(* IEC 61131-3 sources: plc-st-coding-agent/progress/evidence/f14_v14_remaining_20261113/jobs/codex_minimax-m27 (part 4) *)

(* ---- public-medium-04.patch_base_04.st ---- *)
FUNCTION_BLOCK FB_TemperatureControl
VAR_INPUT
    TemperatureSensorInput : REAL;
    SetTemperature : REAL;
END_VAR

VAR_OUTPUT
    CurrentTemperature : REAL;
    SetTempDisplay : REAL;
    HeaterStatus : BOOL;
    OverheatProtection : BOOL;
    HeaterOutput : BOOL;
END_VAR

VAR
    HeaterRuntimeTimer : TON;
    OverheatCooldownTimer : TON;
    tmp_InOverheatProtection : BOOL;
    tmp_SensorFault : BOOL;
    tmp_HeaterShouldBeOn : BOOL;
END_VAR

(*
ENGINEERING_CONTRACT
================================================================================
| Output/State        | Activation          | Retention/Reset           | Units/Boundaries     |
|---------------------|---------------------|---------------------------|----------------------|
| CurrentTemperature  | Every scan (copy)   | Unchanged when fault      | REAL, no conversion  |
| SetTempDisplay      | Every scan (copy)   | Always updated            | REAL, no conversion  |
| HeaterStatus        | Every scan (AND)    | False on fault or overheat| BOOL, same-scan      |
| OverheatProtection  | tmp_InOverheatProt  | Hold 3s cooldown then OFF | BOOL, timer-driven   |
| HeaterOutput        | temp < set && !prot | Off on fault, >5s prot,   | BOOL, 5s threshold   |
|                     |                     |   or temp >= set          | > not >= per spec    |
================================================================================
PUB001: temp < set triggers heater on
PUB002: temp > set turns heater off
PUB003: >5s continuous heater runtime triggers overheat protection
PUB004: 3s cooldown before overheat protection can be lifted
PUB005: Sensor fault if input < 0 or > 100
PUB006: Display current temp, set temp, heater status, overheat status
PUB007: Heater must be off during sensor fault
PUB008: Heater off during overheat protection until cooldown completes
================================================================================

CONTRACT_RULES []
*)

// Update display outputs every scan
CurrentTemperature := TemperatureSensorInput;
SetTempDisplay := SetTemperature;

// Detect sensor fault: temperature out of valid range [0, 100]
tmp_SensorFault := (TemperatureSensorInput < 0.0) OR (TemperatureSensorInput > 100.0);

// Determine if heater should be on (based on temperature comparison only)
tmp_HeaterShouldBeOn := (NOT tmp_SensorFault) AND (TemperatureSensorInput < SetTemperature);

// Overheat protection state machine
IF NOT tmp_InOverheatProtection THEN
    // Normal operation: check if overheat protection should trigger
    IF tmp_HeaterShouldBeOn THEN
        // Heater is on, start accumulating runtime
        HeaterRuntimeTimer(IN := TRUE, PT := T#5S);
        IF HeaterRuntimeTimer.Q THEN
            // Heater ran for more than 5 seconds continuously
            tmp_InOverheatProtection := TRUE;
            HeaterRuntimeTimer(IN := FALSE);
        END_IF;
    ELSE
        // Heater is off, reset runtime timer
        HeaterRuntimeTimer(IN := FALSE);
    END_IF;
ELSE
    // In overheat protection state, start 3-second cooldown
    HeaterRuntimeTimer(IN := FALSE);
    OverheatCooldownTimer(IN := TRUE, PT := T#3S);
    IF OverheatCooldownTimer.Q THEN
        // Cooldown complete, clear overheat protection
        tmp_InOverheatProtection := FALSE;
        OverheatCooldownTimer(IN := FALSE);
    END_IF;
END_IF;

// Update overheat protection output
OverheatProtection := tmp_InOverheatProtection;

// Calculate final heater output
// HeaterOutput is true when:
//   - Temperature is below setpoint
//   - Not in sensor fault
//   - Not in overheat protection
HeaterOutput := tmp_HeaterShouldBeOn AND (NOT tmp_InOverheatProtection);

// Heater status follows actual heater output
HeaterStatus := HeaterOutput;

END_FUNCTION_BLOCK

(* ---- public-medium-04.raw_candidate_01.st ---- *)
FUNCTION_BLOCK FB_TemperatureControl
VAR_INPUT
    TemperatureSensorInput : REAL;
    SetTemperature : REAL;
END_VAR

VAR_OUTPUT
    CurrentTemperature : REAL;
    SetTempDisplay : REAL;
    HeaterStatus : BOOL;
    OverheatProtection : BOOL;
    HeaterOutput : BOOL;
END_VAR

VAR
    HeaterRuntimeTimer : TON;
    OverheatCooldownTimer : TON;
    tmp_InOverheatProtection : BOOL;
    tmp_SensorFault : BOOL;
END_VAR

(*
ENGINEERING_CONTRACT
================================================================================
| Output/State        | Activation          | Retention/Reset           | Units/Boundaries     |
|---------------------|---------------------|---------------------------|----------------------|
| CurrentTemperature  | Every scan (copy)   | Unchanged when fault      | REAL, no conversion  |
| SetTempDisplay      | Every scan (copy)   | Always updated            | REAL, no conversion  |
| HeaterStatus        | Every scan (AND)    | False on fault or overheat| BOOL, same-scan      |
| OverheatProtection  | tmp_InOverheatProt  | Hold 3s cooldown then OFF | BOOL, timer-driven   |
| HeaterOutput        | temp < set && !prot | Off on fault, >5s prot,   | BOOL, 5s threshold   |
|                     |                     |   or temp >= set          | > not >= per spec    |
================================================================================
PUB001: temp < set triggers heater on
PUB002: temp > set turns heater off
PUB003: >5s continuous heater runtime triggers overheat protection
PUB004: 3s cooldown before overheat protection can be lifted
PUB005: Sensor fault if input < 0 or > 100
PUB006: Display current temp, set temp, heater status, overheat status
PUB007: Heater must be off during sensor fault
PUB008: Heater off during overheat protection until cooldown completes
================================================================================

CONTRACT_RULES []
*)

// Update display outputs every scan
CurrentTemperature := TemperatureSensorInput;
SetTempDisplay := SetTemperature;

// Detect sensor fault: temperature out of valid range [0, 100]
tmp_SensorFault := (TemperatureSensorInput < 0.0) OR (TemperatureSensorInput > 100.0);

// Determine if heater should be on (based on temperature comparison only)
tmp_HeaterShouldBeOn := (NOT tmp_SensorFault) AND (TemperatureSensorInput < SetTemperature);

// Overheat protection state machine
IF NOT tmp_InOverheatProtection THEN
    // Normal operation: check if overheat protection should trigger
    IF tmp_HeaterShouldBeOn THEN
        // Heater is on, start accumulating runtime
        HeaterRuntimeTimer(IN := TRUE, PT := T#5S);
        IF HeaterRuntimeTimer.Q THEN
            // Heater ran for more than 5 seconds continuously
            tmp_InOverheatProtection := TRUE;
            HeaterRuntimeTimer(IN := FALSE);
        END_IF;
    ELSE
        // Heater is off, reset runtime timer
        HeaterRuntimeTimer(IN := FALSE);
    END_IF;
ELSE
    // In overheat protection state, start 3-second cooldown
    HeaterRuntimeTimer(IN := FALSE);
    OverheatCooldownTimer(IN := TRUE, PT := T#3S);
    IF OverheatCooldownTimer.Q THEN
        // Cooldown complete, clear overheat protection
        tmp_InOverheatProtection := FALSE;
        OverheatCooldownTimer(IN := FALSE);
    END_IF;
END_IF;

// Update overheat protection output
OverheatProtection := tmp_InOverheatProtection;

// Calculate final heater output
// HeaterOutput is true when:
//   - Temperature is below setpoint
//   - Not in sensor fault
//   - Not in overheat protection
HeaterOutput := tmp_HeaterShouldBeOn AND (NOT tmp_InOverheatProtection);

// Heater status follows actual heater output
HeaterStatus := HeaterOutput;

END_FUNCTION_BLOCK

(* ---- public-medium-04.raw_candidate_02.st ---- *)
FUNCTION_BLOCK FB_TemperatureControl
VAR_INPUT
    TemperatureSensorInput : REAL;
    SetTemperature : REAL;
END_VAR

VAR_OUTPUT
    CurrentTemperature : REAL;
    SetTempDisplay : REAL;
    HeaterStatus : BOOL;
    OverheatProtection : BOOL;
    HeaterOutput : BOOL;
END_VAR

VAR
    HeaterRuntimeTimer : TON;
    OverheatCooldownTimer : TON;
    tmp_InOverheatProtection : BOOL;
    tmp_SensorFault : BOOL;
    tmp_HeaterShouldBeOn : BOOL;
END_VAR

(*
ENGINEERING_CONTRACT
================================================================================
| Output/State        | Activation          | Retention/Reset           | Units/Boundaries     |
|---------------------|---------------------|---------------------------|----------------------|
| CurrentTemperature  | Every scan (copy)   | Unchanged when fault      | REAL, no conversion  |
| SetTempDisplay      | Every scan (copy)   | Always updated            | REAL, no conversion  |
| HeaterStatus        | Every scan (AND)    | False on fault or overheat| BOOL, same-scan      |
| OverheatProtection  | tmp_InOverheatProt  | Hold 3s cooldown then OFF | BOOL, timer-driven   |
| HeaterOutput        | temp < set && !prot | Off on fault, >5s prot,   | BOOL, 5s threshold   |
|                     |                     |   or temp >= set          | > not >= per spec    |
================================================================================
PUB001: temp < set triggers heater on
PUB002: temp > set turns heater off
PUB003: >5s continuous heater runtime triggers overheat protection
PUB004: 3s cooldown before overheat protection can be lifted
PUB005: Sensor fault if input < 0 or > 100
PUB006: Display current temp, set temp, heater status, overheat status
PUB007: Heater must be off during sensor fault
PUB008: Heater off during overheat protection until cooldown completes
================================================================================

CONTRACT_RULES []
*)

// Update display outputs every scan
CurrentTemperature := TemperatureSensorInput;
SetTempDisplay := SetTemperature;

// Detect sensor fault: temperature out of valid range [0, 100]
tmp_SensorFault := (TemperatureSensorInput < 0.0) OR (TemperatureSensorInput > 100.0);

// Determine if heater should be on (based on temperature comparison only)
tmp_HeaterShouldBeOn := (NOT tmp_SensorFault) AND (TemperatureSensorInput < SetTemperature);

// Overheat protection state machine
IF NOT tmp_InOverheatProtection THEN
    // Normal operation: check if overheat protection should trigger
    IF tmp_HeaterShouldBeOn THEN
        // Heater is on, start accumulating runtime
        HeaterRuntimeTimer(IN := TRUE, PT := T#5S);
        IF HeaterRuntimeTimer.Q THEN
            // Heater ran for more than 5 seconds continuously
            tmp_InOverheatProtection := TRUE;
            HeaterRuntimeTimer(IN := FALSE);
        END_IF;
    ELSE
        // Heater is off, reset runtime timer
        HeaterRuntimeTimer(IN := FALSE);
    END_IF;
ELSE
    // In overheat protection state, start 3-second cooldown
    HeaterRuntimeTimer(IN := FALSE);
    OverheatCooldownTimer(IN := TRUE, PT := T#3S);
    IF OverheatCooldownTimer.Q THEN
        // Cooldown complete, clear overheat protection
        tmp_InOverheatProtection := FALSE;
        OverheatCooldownTimer(IN := FALSE);
    END_IF;
END_IF;

// Update overheat protection output
OverheatProtection := tmp_InOverheatProtection;

// Calculate final heater output
// HeaterOutput is true when:
//   - Temperature is below setpoint
//   - Not in sensor fault
//   - Not in overheat protection
HeaterOutput := tmp_HeaterShouldBeOn AND (NOT tmp_InOverheatProtection);

// Heater status follows actual heater output
HeaterStatus := HeaterOutput;

END_FUNCTION_BLOCK

(* ---- public-medium-04.raw_candidate_04.st ---- *)
FUNCTION_BLOCK FB_TemperatureControl
VAR_INPUT
    TemperatureSensorInput : REAL;
    SetTemperature : REAL;
END_VAR

VAR_OUTPUT
    CurrentTemperature : REAL;
    SetTempDisplay : REAL;
    HeaterStatus : BOOL;
    OverheatProtection : BOOL;
    HeaterOutput : BOOL;
END_VAR

VAR
    HeaterRuntimeTimer : TON;
    OverheatCooldownTimer : TON;
    tmp_InOverheatProtection : BOOL;
    tmp_SensorFault : BOOL;
    tmp_RuntimeTimerEnable : BOOL;
END_VAR

(*
ENGINEERING_CONTRACT
================================================================================
| Output/State        | Activation          | Retention/Reset           | Units/Boundaries     |
|---------------------|---------------------|---------------------------|----------------------|
| CurrentTemperature  | Every scan (copy)   | Unchanged when fault      | REAL, no conversion  |
| SetTempDisplay      | Every scan (copy)   | Always updated            | REAL, no conversion  |
| HeaterStatus        | Every scan (AND)    | False on fault or overheat| BOOL, same-scan      |
| OverheatProtection  | tmp_InOverheatProt  | Hold 3s cooldown then OFF | BOOL, timer-driven   |
| HeaterOutput        | temp < set && !prot | Off on fault, >5s prot,   | BOOL, 5s threshold   |
|                     |                     |   or temp >= set          | > not >= per spec    |
================================================================================
PUB001: temp < set triggers heater on
PUB002: temp > set turns heater off
PUB003: >5s continuous heater runtime triggers overheat protection
PUB004: 3s cooldown before overheat protection can be lifted
PUB005: Sensor fault if input < 0 or > 100
PUB006: Display current temp, set temp, heater status, overheat status
PUB007: Heater must be off during sensor fault
PUB008: Heater off during overheat protection until cooldown completes
================================================================================

CONTRACT_RULES []
*)

// Update display outputs every scan
CurrentTemperature := TemperatureSensorInput;
SetTempDisplay := SetTemperature;

// Detect sensor fault: temperature out of valid range [0, 100]
tmp_SensorFault := (TemperatureSensorInput < 0.0) OR (TemperatureSensorInput > 100.0);

// Determine if runtime timer should accumulate (heater on, not in fault, not in overheat protection)
tmp_RuntimeTimerEnable := (NOT tmp_SensorFault) AND (NOT tmp_InOverheatProtection) AND (TemperatureSensorInput < SetTemperature);

// Overheat protection state machine
IF NOT tmp_InOverheatProtection THEN
    // Normal operation: check if overheat protection should trigger
    IF tmp_RuntimeTimerEnable THEN
        // Heater is on, start accumulating runtime
        HeaterRuntimeTimer(IN := TRUE, PT := T#5001MS);
        IF HeaterRuntimeTimer.Q THEN
            // Heater ran for more than 5 seconds continuously
            tmp_InOverheatProtection := TRUE;
            HeaterRuntimeTimer(IN := FALSE);
        END_IF;
    ELSE
        // Heater is off or in fault, reset runtime timer
        HeaterRuntimeTimer(IN := FALSE);
    END_IF;
ELSE
    // In overheat protection state, run 3-second cooldown
    HeaterRuntimeTimer(IN := FALSE);
    OverheatCooldownTimer(IN := TRUE, PT := T#3S);
    IF OverheatCooldownTimer.Q THEN
        // Cooldown complete, clear overheat protection
        tmp_InOverheatProtection := FALSE;
        OverheatCooldownTimer(IN := FALSE);
    END_IF;
END_IF;

// Update outputs
OverheatProtection := tmp_InOverheatProtection;

// Calculate final heater output: on when temperature below setpoint, not in fault, not in overheat protection
HeaterOutput := tmp_RuntimeTimerEnable;

// Heater status follows actual heater output
HeaterStatus := HeaterOutput;

END_FUNCTION_BLOCK

(* ---- public-medium-05.candidate_01.st ---- *)
(* ENGINEERING_CONTRACT *)
(*
Mode behavior (PUB001):
- Mode=0: Manual mode (ForwardButton→MotorForward, ReverseButton→MotorReverse)
- Mode=1: Automatic mode (A→B→C state machine)

Manual mode (PUB002):
- MotorForward activates with ForwardButton when Mode=0, interlocked with ReverseButton
- MotorReverse activates with ReverseButton when Mode=0, interlocked with ForwardButton
- CompletionLight always OFF in manual mode

Automatic mode (PUB003):
- IDLE→SensorA: wait at Station A for ButtonA press
- Station A: MotorForward TRUE while State=MOVING_TO_B
- MOVING_TO_B→SensorB: hold at Station B for ButtonB press
- Station B: MotorForward TRUE while State=MOVING_TO_C
- MOVING_TO_C→SensorC: hold at Station C

CompletionLight behavior (PUB006, PUB007, PUB008):
- Activation: State=STATION_C AND SensorC AND ButtonC (same-scan)
- Retention: State=STATION_C AND SensorC (CompletionLight remains TRUE)
- Deactivation: State≠STATION_C OR NOT SensorC (product removal)
- Units: boolean, no units

Output states:
- MotorForward: combinational in manual, pulsed in auto (A→B, B→C transitions)
- MotorReverse: combinational in manual only, always FALSE in auto
- CompletionLight: retained while product at Station C, no explicit reset input

Scan priority: same-scan evaluation of all conditions before outputs
*)

(* CONTRACT_RULES [] *)

FUNCTION_BLOCK ProductionLineControl
VAR_INPUT
    Mode            : BOOL;
    ForwardButton   : BOOL;
    ReverseButton   : BOOL;
    SensorA         : BOOL;
    SensorB         : BOOL;
    SensorC         : BOOL;
    ButtonA         : BOOL;
    ButtonB         : BOOL;
    ButtonC         : BOOL;
END_VAR
VAR_OUTPUT
    MotorForward    : BOOL;
    MotorReverse    : BOOL;
    CompletionLight : BOOL;
END_VAR
VAR
    State : INT;
END_VAR

// State constants
CONSTANTS
    STATE_IDLE         : INT := 0;
    STATE_STATION_A    : INT := 1;
    STATE_MOVING_TO_B  : INT := 2;
    STATE_STATION_B    : INT := 3;
    STATE_MOVING_TO_C  : INT := 4;
    STATE_STATION_C    : INT := 5;
END_CONSTANTS

// Initialize state on first call
IF State = 0 THEN
    State := STATE_IDLE;
END_IF;

// Manual mode: direct button control with direction interlock
IF Mode = FALSE THEN
    MotorForward := ForwardButton AND NOT ReverseButton;
    MotorReverse := ReverseButton AND NOT ForwardButton;
    CompletionLight := FALSE;
    State := STATE_IDLE;
ELSE
    // Automatic mode: state machine control
    IF State = STATE_IDLE THEN
        MotorForward := FALSE;
        MotorReverse := FALSE;
        CompletionLight := FALSE;

        IF SensorA THEN
            State := STATE_STATION_A;
        END_IF;

    ELSIF State = STATE_STATION_A THEN
        MotorForward := FALSE;

        IF ButtonA THEN
            State := STATE_MOVING_TO_B;
        END_IF;

    ELSIF State = STATE_MOVING_TO_B THEN
        MotorForward := TRUE;

        IF SensorB THEN
            MotorForward := FALSE;
            State := STATE_STATION_B;
        END_IF;

    ELSIF State = STATE_STATION_B THEN
        MotorForward := FALSE;

        IF ButtonB THEN
            State := STATE_MOVING_TO_C;
        END_IF;

    ELSIF State = STATE_MOVING_TO_C THEN
        MotorForward := TRUE;

        IF SensorC THEN
            MotorForward := FALSE;
            State := STATE_STATION_C;
        END_IF;

    ELSIF State = STATE_STATION_C THEN
        MotorForward := FALSE;

        IF NOT SensorC THEN
            State := STATE_IDLE;
            CompletionLight := FALSE;
        ELSE
            CompletionLight := TRUE;
        END_IF;
    END_IF;
END_IF;

END_FUNCTION_BLOCK

(* ---- public-medium-05.patch_base_02.st ---- *)
(* ENGINEERING_CONTRACT *)
(*
Mode behavior (PUB001):
- Mode=0: Manual mode (ForwardButton→MotorForward, ReverseButton→MotorReverse)
- Mode=1: Automatic mode (A→B→C state machine)

Manual mode (PUB002):
- MotorForward activates with ForwardButton when Mode=0, interlocked with ReverseButton
- MotorReverse activates with ReverseButton when Mode=0, interlocked with ForwardButton
- CompletionLight always OFF in manual mode

Automatic mode (PUB003):
- IDLE→SensorA: wait at Station A for ButtonA press
- Station A: MotorForward TRUE while State=MOVING_TO_B
- MOVING_TO_B→SensorB: hold at Station B for ButtonB press
- Station B: MotorForward TRUE while State=MOVING_TO_C
- MOVING_TO_C→SensorC: hold at Station C

CompletionLight behavior (PUB006, PUB007, PUB008):
- Activation: State=STATION_C AND SensorC AND ButtonC (same-scan)
- Retention: State=STATION_C AND SensorC (CompletionLight remains TRUE)
- Deactivation: State≠STATION_C OR NOT SensorC (product removal)
- Units: boolean, no units

Output states:
- MotorForward: combinational in manual, pulsed in auto (A→B, B→C transitions)
- MotorReverse: combinational in manual only, always FALSE in auto
- CompletionLight: retained while product at Station C, no explicit reset input

Scan priority: same-scan evaluation of all conditions before outputs
*)

(* CONTRACT_RULES [] *)

FUNCTION_BLOCK ProductionLineControl
VAR_INPUT
    Mode            : BOOL;
    ForwardButton   : BOOL;
    ReverseButton   : BOOL;
    SensorA         : BOOL;
    SensorB         : BOOL;
    SensorC         : BOOL;
    ButtonA         : BOOL;
    ButtonB         : BOOL;
    ButtonC         : BOOL;
END_VAR
VAR_OUTPUT
    MotorForward    : BOOL;
    MotorReverse    : BOOL;
    CompletionLight : BOOL;
END_VAR
VAR
    State : INT;
END_VAR

// State constants
CONSTANTS
    STATE_IDLE         : INT := 0;
    STATE_STATION_A    : INT := 1;
    STATE_MOVING_TO_B  : INT := 2;
    STATE_STATION_B    : INT := 3;
    STATE_MOVING_TO_C  : INT := 4;
    STATE_STATION_C    : INT := 5;
END_CONSTANTS

// Initialize state on first call
IF State = 0 THEN
    State := STATE_IDLE;
END_IF;

// Manual mode: direct button control with direction interlock
IF Mode = FALSE THEN
    MotorForward := ForwardButton AND NOT ReverseButton;
    MotorReverse := ReverseButton AND NOT ForwardButton;
    CompletionLight := FALSE;
    State := STATE_IDLE;
ELSE
    // Automatic mode: state machine control
    IF State = STATE_IDLE THEN
        MotorForward := FALSE;
        MotorReverse := FALSE;
        CompletionLight := FALSE;

        IF SensorA THEN
            State := STATE_STATION_A;
        END_IF;

    ELSIF State = STATE_STATION_A THEN
        MotorForward := FALSE;

        IF ButtonA THEN
            State := STATE_MOVING_TO_B;
        END_IF;

    ELSIF State = STATE_MOVING_TO_B THEN
        MotorForward := TRUE;

        IF SensorB THEN
            MotorForward := FALSE;
            State := STATE_STATION_B;
        END_IF;

    ELSIF State = STATE_STATION_B THEN
        MotorForward := FALSE;

        IF ButtonB THEN
            State := STATE_MOVING_TO_C;
        END_IF;

    ELSIF State = STATE_MOVING_TO_C THEN
        MotorForward := TRUE;

        IF SensorC THEN
            MotorForward := FALSE;
            State := STATE_STATION_C;
        END_IF;

    ELSIF State = STATE_STATION_C THEN
        MotorForward := FALSE;

        IF NOT SensorC THEN
            State := STATE_IDLE;
            CompletionLight := FALSE;
        ELSE
            CompletionLight := TRUE;
        END_IF;
    END_IF;
END_IF;

END_FUNCTION_BLOCK

(* ---- public-medium-05.patch_base_03.st ---- *)
(* ENGINEERING_CONTRACT *)
(*
Mode behavior (PUB001):
- Mode=0: Manual mode (ForwardButton→MotorForward, ReverseButton→MotorReverse)
- Mode=1: Automatic mode (A→B→C state machine)

Manual mode (PUB002):
- MotorForward activates with ForwardButton when Mode=0, interlocked with ReverseButton
- MotorReverse activates with ReverseButton when Mode=0, interlocked with ForwardButton
- CompletionLight always OFF in manual mode

Automatic mode (PUB003):
- IDLE→SensorA: wait at Station A for ButtonA press
- Station A: MotorForward TRUE while State=MOVING_TO_B
- MOVING_TO_B→SensorB: hold at Station B for ButtonB press
- Station B: MotorForward TRUE while State=MOVING_TO_C
- MOVING_TO_C→SensorC: hold at Station C

CompletionLight behavior (PUB006, PUB007, PUB008):
- Activation: State=STATION_C AND SensorC AND ButtonC (same-scan)
- Retention: State=STATION_C AND SensorC (CompletionLight remains TRUE)
- Deactivation: State≠STATION_C OR NOT SensorC (product removal)
- Units: boolean, no units

Output states:
- MotorForward: combinational in manual, pulsed in auto (A→B, B→C transitions)
- MotorReverse: combinational in manual only, always FALSE in auto
- CompletionLight: retained while product at Station C, no explicit reset input

Scan priority: same-scan evaluation of all conditions before outputs
*)

(* CONTRACT_RULES [] *)

FUNCTION_BLOCK ProductionLineControl
VAR_INPUT
    Mode            : BOOL;
    ForwardButton   : BOOL;
    ReverseButton   : BOOL;
    SensorA         : BOOL;
    SensorB         : BOOL;
    SensorC         : BOOL;
    ButtonA         : BOOL;
    ButtonB         : BOOL;
    ButtonC         : BOOL;
END_VAR
VAR_OUTPUT
    MotorForward    : BOOL;
    MotorReverse    : BOOL;
    CompletionLight : BOOL;
END_VAR
VAR
    State : INT;
END_VAR

// State constants
CONSTANTS
    STATE_IDLE         : INT := 0;
    STATE_STATION_A    : INT := 1;
    STATE_MOVING_TO_B  : INT := 2;
    STATE_STATION_B    : INT := 3;
    STATE_MOVING_TO_C  : INT := 4;
    STATE_STATION_C    : INT := 5;
END_CONSTANTS

// Initialize state on first call
IF State = 0 THEN
    State := STATE_IDLE;
END_IF;

// Manual mode: direct button control with direction interlock
IF Mode = FALSE THEN
    MotorForward := ForwardButton AND NOT ReverseButton;
    MotorReverse := ReverseButton AND NOT ForwardButton;
    CompletionLight := FALSE;
    State := STATE_IDLE;
ELSE
    // Automatic mode: state machine control
    IF State = STATE_IDLE THEN
        MotorForward := FALSE;
        MotorReverse := FALSE;
        CompletionLight := FALSE;

        IF SensorA THEN
            State := STATE_STATION_A;
        END_IF;

    ELSIF State = STATE_STATION_A THEN
        MotorForward := FALSE;

        IF ButtonA THEN
            State := STATE_MOVING_TO_B;
        END_IF;

    ELSIF State = STATE_MOVING_TO_B THEN
        MotorForward := TRUE;

        IF SensorB THEN
            MotorForward := FALSE;
            State := STATE_STATION_B;
        END_IF;

    ELSIF State = STATE_STATION_B THEN
        MotorForward := FALSE;

        IF ButtonB THEN
            State := STATE_MOVING_TO_C;
        END_IF;

    ELSIF State = STATE_MOVING_TO_C THEN
        MotorForward := TRUE;

        IF SensorC THEN
            MotorForward := FALSE;
            State := STATE_STATION_C;
        END_IF;

    ELSIF State = STATE_STATION_C THEN
        MotorForward := FALSE;

        IF NOT SensorC THEN
            State := STATE_IDLE;
            CompletionLight := FALSE;
        ELSE
            CompletionLight := TRUE;
        END_IF;
    END_IF;
END_IF;

END_FUNCTION_BLOCK

(* ---- public-medium-05.raw_candidate_01.st ---- *)
(* ENGINEERING_CONTRACT *)
(*
Mode behavior (PUB001):
- Mode=0: Manual mode (ForwardButton→MotorForward, ReverseButton→MotorReverse)
- Mode=1: Automatic mode (A→B→C state machine)

Manual mode (PUB002):
- MotorForward activates with ForwardButton when Mode=0, interlocked with ReverseButton
- MotorReverse activates with ReverseButton when Mode=0, interlocked with ForwardButton
- CompletionLight always OFF in manual mode

Automatic mode (PUB003):
- IDLE→SensorA: wait at Station A for ButtonA press
- Station A: MotorForward TRUE while State=MOVING_TO_B
- MOVING_TO_B→SensorB: hold at Station B for ButtonB press
- Station B: MotorForward TRUE while State=MOVING_TO_C
- MOVING_TO_C→SensorC: hold at Station C

CompletionLight behavior (PUB006, PUB007, PUB008):
- Activation: State=STATION_C AND SensorC AND ButtonC (same-scan)
- Retention: State=STATION_C AND SensorC (CompletionLight remains TRUE)
- Deactivation: State≠STATION_C OR NOT SensorC (product removal)
- Units: boolean, no units

Output states:
- MotorForward: combinational in manual, pulsed in auto (A→B, B→C transitions)
- MotorReverse: combinational in manual only, always FALSE in auto
- CompletionLight: retained while product at Station C, no explicit reset input

Scan priority: same-scan evaluation of all conditions before outputs
*)

(* CONTRACT_RULES [] *)

FUNCTION_BLOCK ProductionLineControl
VAR_INPUT
    Mode            : BOOL;
    ForwardButton   : BOOL;
    ReverseButton   : BOOL;
    SensorA         : BOOL;
    SensorB         : BOOL;
    SensorC         : BOOL;
    ButtonA         : BOOL;
    ButtonB         : BOOL;
    ButtonC         : BOOL;
END_VAR
VAR_OUTPUT
    MotorForward    : BOOL;
    MotorReverse    : BOOL;
    CompletionLight : BOOL;
END_VAR
VAR
    State : INT;
END_VAR

// State constants
CONSTANTS
    STATE_IDLE         : INT := 0;
    STATE_STATION_A    : INT := 1;
    STATE_MOVING_TO_B  : INT := 2;
    STATE_STATION_B    : INT := 3;
    STATE_MOVING_TO_C  : INT := 4;
    STATE_STATION_C    : INT := 5;
END_CONSTANTS

// Initialize state on first call
IF State = 0 THEN
    State := STATE_IDLE;
END_IF

// Manual mode: direct button control with direction interlock
IF Mode = FALSE THEN
    MotorForward := ForwardButton AND NOT ReverseButton;
    MotorReverse := ReverseButton AND NOT ForwardButton;
    CompletionLight := FALSE;
    State := STATE_IDLE;
ELSE
    // Automatic mode: state machine control
    IF State = STATE_IDLE THEN
        MotorForward := FALSE;
        MotorReverse := FALSE;
        CompletionLight := FALSE;

        IF SensorA THEN
            State := STATE_STATION_A;
        END_IF

    ELSIF State = STATE_STATION_A THEN
        MotorForward := FALSE;

        IF ButtonA THEN
            State := STATE_MOVING_TO_B;
        END_IF

    ELSIF State = STATE_MOVING_TO_B THEN
        MotorForward := TRUE;

        IF SensorB THEN
            MotorForward := FALSE;
            State := STATE_STATION_B;
        END_IF

    ELSIF State = STATE_STATION_B THEN
        MotorForward := FALSE;

        IF ButtonB THEN
            State := STATE_MOVING_TO_C;
        END_IF

    ELSIF State = STATE_MOVING_TO_C THEN
        MotorForward := TRUE;

        IF SensorC THEN
            MotorForward := FALSE;
            State := STATE_STATION_C;
        END_IF

    ELSIF State = STATE_STATION_C THEN
        MotorForward := FALSE;

        IF NOT SensorC THEN
            State := STATE_IDLE;
            CompletionLight := FALSE;
        ELSE
            CompletionLight := TRUE;
        END_IF
    END_IF
END_IF

END_FUNCTION_BLOCK

(* ---- public-medium-06.candidate_01.st ---- *)
FUNCTION_BLOCK SlabThicknessMonitor
VAR_INPUT
    THICKNESS_FAULT        : BOOL;
    THICKNESS_SIGNAL_VALID : BOOL;
    CUTTING_RUN            : BOOL;
    FaultTimestamp         : DINT;
    CycleTime              : TIME;
END_VAR

VAR_OUTPUT
    THICKNESS_ALARM           : BOOL := FALSE;
    Slab_Fault_Counter        : UINT := 0;
    Slab_Runtime_Accumulator  : LTIME := LTIME#0s;
    Slab_Fault_History        : ARRAY[0..4] OF DINT := [5(0)];
END_VAR

VAR
    tmp_AlarmHoldTimer : TON;
    tmp_FaultRTrig     : R_TRIG;
END_VAR

(*
ENGINEERING_CONTRACT
================================================================================
| Output / State        | Activation              | Retention/Reset            |
|-----------------------|-------------------------|----------------------------|
| THICKNESS_ALARM       | Rising edge valid fault | Reset: signal invalid/Power|
| Hold Timer (500ms)    | Rising edge valid fault | Reset: elapsed or invalid  |
| Slab_Fault_Counter    | Rising edge valid fault | Retention: no reset        |
| Slab_Fault_History[0] | Rising edge valid fault | Shift register, newest=0   |
| Slab_Runtime_Accum.   | CUTTING_RUN+valid+no    | Retention: preserve unless |
|                       | fault per scan          | condition met              |
--------------------------------------------------------------------------------
Priority: Same-scan; alarm combinational with hold timer; no edge-only reset.
Units: LTIME nanoseconds; CycleTime T#1ms..T#1h; hold = T#500ms >= 500ms.
Boundaries: History array fixed 0..4; counter saturates at UINT MAX.
Pub Refs: PUB001, PUB002, PUB003, PUB004, PUB005, PUB006
================================================================================
*)

(* CONTRACT_RULES [] *)

tmp_FaultRTrig(CLK := THICKNESS_FAULT AND THICKNESS_SIGNAL_VALID);

IF tmp_FaultRTrig.Q THEN
    tmp_AlarmHoldTimer(IN := TRUE, PT := T#500ms);
END_IF;

IF tmp_AlarmHoldTimer.Q THEN
    tmp_AlarmHoldTimer(IN := FALSE);
END_IF;

IF NOT THICKNESS_SIGNAL_VALID THEN
    THICKNESS_ALARM := FALSE;
    tmp_AlarmHoldTimer(IN := FALSE);
ELSIF THICKNESS_FAULT THEN
    THICKNESS_ALARM := TRUE;
    tmp_AlarmHoldTimer(IN := TRUE, PT := T#500ms);
ELSIF tmp_AlarmHoldTimer.Q THEN
    THICKNESS_ALARM := TRUE;
ELSE
    THICKNESS_ALARM := FALSE;
END_IF;

IF CUTTING_RUN AND THICKNESS_SIGNAL_VALID AND NOT THICKNESS_FAULT THEN
    Slab_Runtime_Accumulator := Slab_Runtime_Accumulator + TO_LTIME(CycleTime);
END_IF;

IF tmp_FaultRTrig.Q THEN
    Slab_Fault_History[4] := Slab_Fault_History[3];
    Slab_Fault_History[3] := Slab_Fault_History[2];
    Slab_Fault_History[2] := Slab_Fault_History[1];
    Slab_Fault_History[1] := Slab_Fault_History[0];
    Slab_Fault_History[0] := FaultTimestamp;
    Slab_Fault_Counter := Slab_Fault_Counter + UINT#1;
END_IF;

END_FUNCTION_BLOCK

(* ---- public-medium-06.raw_candidate_01.st ---- *)
FUNCTION_BLOCK SlabThicknessMonitor
VAR_INPUT
    THICKNESS_FAULT        : BOOL;
    THICKNESS_SIGNAL_VALID : BOOL;
    CUTTING_RUN            : BOOL;
    FaultTimestamp         : DINT;
    CycleTime              : TIME;
END_VAR

VAR_OUTPUT
    THICKNESS_ALARM           : BOOL := FALSE;
    Slab_Fault_Counter        : UINT := 0;
    Slab_Runtime_Accumulator  : LTIME := LTIME#0s;
    Slab_Fault_History        : ARRAY[0..4] OF DINT := [5(0)];
END_VAR

VAR
    tmp_AlarmHoldTimer : TON;
    tmp_FaultRTrig     : R_TRIG;
END_VAR

(*
ENGINEERING_CONTRACT
================================================================================
| Output / State        | Activation              | Retention/Reset            |
|-----------------------|-------------------------|----------------------------|
| THICKNESS_ALARM       | Rising edge valid fault | Reset: signal invalid/Power|
| Hold Timer (500ms)    | Rising edge valid fault | Reset: elapsed or invalid  |
| Slab_Fault_Counter    | Rising edge valid fault | Retention: no reset        |
| Slab_Fault_History[0] | Rising edge valid fault | Shift register, newest=0   |
| Slab_Runtime_Accum.   | CUTTING_RUN+valid+no    | Retention: preserve unless |
|                       | fault per scan          | condition met              |
--------------------------------------------------------------------------------
Priority: Same-scan; alarm combinational with hold timer; no edge-only reset.
Units: LTIME nanoseconds; CycleTime T#1ms..T#1h; hold = T#500ms >= 500ms.
Boundaries: History array fixed 0..4; counter saturates at UINT MAX.
Pub Refs: PUB001, PUB002, PUB003, PUB004, PUB005, PUB006
================================================================================
*)

(* CONTRACT_RULES [] *)

tmp_FaultRTrig(CLK := THICKNESS_FAULT AND THICKNESS_SIGNAL_VALID);

IF tmp_FaultRTrig.Q THEN
    tmp_AlarmHoldTimer(IN := TRUE, PT := T#500ms);
END_IF;

IF tmp_AlarmHoldTimer.Q THEN
    tmp_AlarmHoldTimer(IN := FALSE);
END_IF;

IF NOT THICKNESS_SIGNAL_VALID THEN
    THICKNESS_ALARM := FALSE;
    tmp_AlarmHoldTimer(IN := FALSE);
ELSIF THICKNESS_FAULT THEN
    THICKNESS_ALARM := TRUE;
    tmp_AlarmHoldTimer(IN := TRUE, PT := T#500ms);
ELSIF tmp_AlarmHoldTimer.Q THEN
    THICKNESS_ALARM := TRUE;
ELSE
    THICKNESS_ALARM := FALSE;
END_IF;

IF CUTTING_RUN AND THICKNESS_SIGNAL_VALID AND NOT THICKNESS_FAULT THEN
    Slab_Runtime_Accumulator := Slab_Runtime_Accumulator + TO_LTIME(CycleTime);
END_IF;

IF tmp_FaultRTrig.Q THEN
    Slab_Fault_History[4] := Slab_Fault_History[3];
    Slab_Fault_History[3] := Slab_Fault_History[2];
    Slab_Fault_History[2] := Slab_Fault_History[1];
    Slab_Fault_History[1] := Slab_Fault_History[0];
    Slab_Fault_History[0] := FaultTimestamp;
    Slab_Fault_Counter := Slab_Fault_Counter + UINT#1;
END_IF;

END_FUNCTION_BLOCK

(* ---- public-medium-07.candidate_01.st ---- *)
FUNCTION_BLOCK HVAC_Control
(*
ENGINEERING_CONTRACT
| Output/State      | Activation              | Retention           | Reset/Deactivation        | Priority   | Units/Bounds       |
|-------------------|-------------------------|---------------------|---------------------------|------------|--------------------|
| SUPPLY_FAN_RUN    | Occupied + Non-Night,   | Hold while cond met | Unoccupied OR Night mode  | Same-scan  | 30s delay (LTIME)  |
|                   | after 30s TON.Q         |                     | resets TON, stops fan     |            |                    |
| TEMP_SETPOINT_    | Every scan from         | Hold last computed  | Re-evaluated each scan    | Same-scan  | INT ±4°C           |
| ADJUST            | HVAC_MODE_SELECTOR +    | value               | based on mode+occupancy   |            |                    |
|                   | OCCUPANCY_DETECTED +    |                     |                           |            |                    |
|                   | ENERGY_SAVING_MODE      |                     |                           |            |                    |
PUB001: Start 30s delay when OCCUPANCY_DETECTED AND HVAC_MODE_SELECTOR<>3
PUB002: Reset timer and stop fan if OCCUPANCY_DETECTED=FALSE OR HVAC_MODE_SELECTOR=3
PUB003: Temp adj: Auto(0°occ, +3°unocc_ES, +2°unocc_std), Comfort(0°occ, +1°unocc), Economy(0°occ, +4°unocc)
PUB004: Night: +4°C regardless of occupancy
PUB005: ENERGY_SAVING_MODE affects Auto mode only
PUB006: TEMP_SETPOINT_ADJUST within ±4°C
PUB007: Initialize outputs OFF/zero at power-up; update from current inputs
PUB008: Fan start delay controls only BOOL fan enable; no speed ramp
*)
VAR_INPUT
    OCCUPANCY_DETECTED  : BOOL;
    ENERGY_SAVING_MODE  : BOOL;
    HVAC_MODE_SELECTOR  : INT;
END_VAR

VAR_OUTPUT
    SUPPLY_FAN_RUN        : BOOL := FALSE;
    TEMP_SETPOINT_ADJUST  : INT := 0;
END_VAR

VAR
    fanTimer : TON;
END_VAR

// Fan control with 30-second start delay (PUB001, PUB002)
fanTimer(IN := OCCUPANCY_DETECTED AND (HVAC_MODE_SELECTOR <> 3), PT := T#30s);
IF fanTimer.Q THEN
    SUPPLY_FAN_RUN := TRUE;
ELSE
    SUPPLY_FAN_RUN := FALSE;
END_IF;

// Temperature setpoint adjustment (PUB003, PUB004, PUB005, PUB006)
CASE HVAC_MODE_SELECTOR OF
    0: // Auto
        IF OCCUPANCY_DETECTED THEN
            TEMP_SETPOINT_ADJUST := 0;
        ELSE
            IF ENERGY_SAVING_MODE THEN
                TEMP_SETPOINT_ADJUST := 3;
            ELSE
                TEMP_SETPOINT_ADJUST := 2;
            END_IF;
        END_IF;
    1: // Comfort
        IF OCCUPANCY_DETECTED THEN
            TEMP_SETPOINT_ADJUST := 0;
        ELSE
            TEMP_SETPOINT_ADJUST := 1;
        END_IF;
    2: // Economy
        IF OCCUPANCY_DETECTED THEN
            TEMP_SETPOINT_ADJUST := 0;
        ELSE
            TEMP_SETPOINT_ADJUST := 4;
        END_IF;
    3: // Night
        TEMP_SETPOINT_ADJUST := 4;
END_CASE;

// Clamp to ±4°C boundary (PUB006)
IF TEMP_SETPOINT_ADJUST > 4 THEN TEMP_SETPOINT_ADJUST := 4; END_IF;
IF TEMP_SETPOINT_ADJUST < -4 THEN TEMP_SETPOINT_ADJUST := -4; END_IF;

END_FUNCTION_BLOCK

(* ---- public-medium-07.raw_candidate_01.st ---- *)
FUNCTION_BLOCK HVAC_Control
(*
ENGINEERING_CONTRACT
| Output/State      | Activation              | Retention           | Reset/Deactivation        | Priority   | Units/Bounds       |
|-------------------|-------------------------|---------------------|---------------------------|------------|--------------------|
| SUPPLY_FAN_RUN    | Occupied + Non-Night,   | Hold while cond met | Unoccupied OR Night mode  | Same-scan  | 30s delay (LTIME)  |
|                   | after 30s TON.Q         |                     | resets TON, stops fan     |            |                    |
| TEMP_SETPOINT_    | Every scan from         | Hold last computed  | Re-evaluated each scan    | Same-scan  | INT ±4°C           |
| ADJUST            | HVAC_MODE_SELECTOR +    | value               | based on mode+occupancy   |            |                    |
|                   | OCCUPANCY_DETECTED +    |                     |                           |            |                    |
|                   | ENERGY_SAVING_MODE      |                     |                           |            |                    |
PUB001: Start 30s delay when OCCUPANCY_DETECTED AND HVAC_MODE_SELECTOR<>3
PUB002: Reset timer and stop fan if OCCUPANCY_DETECTED=FALSE OR HVAC_MODE_SELECTOR=3
PUB003: Temp adj: Auto(0°occ, +3°unocc_ES, +2°unocc_std), Comfort(0°occ, +1°unocc), Economy(0°occ, +4°unocc)
PUB004: Night: +4°C regardless of occupancy
PUB005: ENERGY_SAVING_MODE affects Auto mode only
PUB006: TEMP_SETPOINT_ADJUST within ±4°C
PUB007: Initialize outputs OFF/zero at power-up; update from current inputs
PUB008: Fan start delay controls only BOOL fan enable; no speed ramp
*)
VAR_INPUT
    OCCUPANCY_DETECTED  : BOOL;
    ENERGY_SAVING_MODE  : BOOL;
    HVAC_MODE_SELECTOR  : INT;
END_VAR

VAR_OUTPUT
    SUPPLY_FAN_RUN        : BOOL := FALSE;
    TEMP_SETPOINT_ADJUST  : INT := 0;
END_VAR

VAR
    fanTimer : TON;
END_VAR

// Fan control with 30-second start delay (PUB001, PUB002)
fanTimer(IN := OCCUPANCY_DETECTED AND (HVAC_MODE_SELECTOR <> 3), PT := T#30s);
IF fanTimer.Q THEN
    SUPPLY_FAN_RUN := TRUE;
ELSE
    SUPPLY_FAN_RUN := FALSE;
END_IF

// Temperature setpoint adjustment (PUB003, PUB004, PUB005, PUB006)
CASE HVAC_MODE_SELECTOR OF
    0: // Auto
        IF OCCUPANCY_DETECTED THEN
            TEMP_SETPOINT_ADJUST := 0;
        ELSE
            IF ENERGY_SAVING_MODE THEN
                TEMP_SETPOINT_ADJUST := 3;
            ELSE
                TEMP_SETPOINT_ADJUST := 2;
            END_IF
        END_IF
    1: // Comfort
        IF OCCUPANCY_DETECTED THEN
            TEMP_SETPOINT_ADJUST := 0;
        ELSE
            TEMP_SETPOINT_ADJUST := 1;
        END_IF
    2: // Economy
        IF OCCUPANCY_DETECTED THEN
            TEMP_SETPOINT_ADJUST := 0;
        ELSE
            TEMP_SETPOINT_ADJUST := 4;
        END_IF
    3: // Night
        TEMP_SETPOINT_ADJUST := 4;
END_CASE

// Clamp to ±4°C boundary (PUB006)
IF TEMP_SETPOINT_ADJUST > 4 THEN TEMP_SETPOINT_ADJUST := 4; END_IF
IF TEMP_SETPOINT_ADJUST < -4 THEN TEMP_SETPOINT_ADJUST := -4; END_IF

END_FUNCTION_BLOCK

(* ---- public-medium-08.candidate_01.st ---- *)
FUNCTION_BLOCK IPv4_Parser
VAR_INPUT
    ipText : STRING(254);
END_VAR
VAR_OUTPUT
    ipValue : UDINT;
END_VAR
VAR
    tmp_pos : UDINT;
    tmp_seg : STRING(4);
    tmp_val : UDINT;
    tmp_byte0 : UDINT;
    tmp_byte1 : UDINT;
    tmp_byte2 : UDINT;
    tmp_byte3 : UDINT;
    tmp_byte_index : UDINT;
    tmp_text_len : UDINT;
    tmp_char : BYTE;
    tmp_seg_len : UDINT;
END_VAR

(*
ENGINEERING_CONTRACT
PUB001: Four nonempty decimal-digit segments separated by periods
PUB002: Each segment 0-255; invalid/empty → ipValue=0
PUB003: Network byte order: seg1=MSB(31:24), seg4=LSB(7:0)
PUB004: Valid address 0.0.0.0 also produces 0 (boundary case)
*)

tmp_text_len := LEN(ipText);
IF tmp_text_len = 0 OR tmp_text_len > 15 THEN
    ipValue := 0;
    RETURN;
END_IF;

tmp_pos := 1;
tmp_byte_index := 0;

WHILE tmp_byte_index < 4 DO
    tmp_seg := '';
    tmp_seg_len := 0;

    WHILE tmp_pos <= tmp_text_len DO
        tmp_char := ipText[tmp_pos - 1];
        IF tmp_char = 46 THEN
            EXIT;
        END_IF;
        IF tmp_char < 48 OR tmp_char > 57 THEN
            ipValue := 0;
            RETURN;
        END_IF;
        tmp_seg := CONCAT(tmp_seg, CHR(tmp_char));
        tmp_seg_len := tmp_seg_len + 1;
        tmp_pos := tmp_pos + 1;
    END_WHILE;

    IF tmp_seg_len = 0 OR tmp_seg_len > 3 THEN
        ipValue := 0;
        RETURN;
    END_IF;

    tmp_val := STRING_TO_UDINT(tmp_seg);
    IF tmp_val > 255 THEN
        ipValue := 0;
        RETURN;
    END_IF;

    IF tmp_byte_index = 0 THEN
        tmp_byte0 := tmp_val;
    ELSIF tmp_byte_index = 1 THEN
        tmp_byte1 := tmp_val;
    ELSIF tmp_byte_index = 2 THEN
        tmp_byte2 := tmp_val;
    ELSIF tmp_byte_index = 3 THEN
        tmp_byte3 := tmp_val;
    END_IF;

    tmp_byte_index := tmp_byte_index + 1;

    IF tmp_pos > tmp_text_len THEN
        EXIT;
    END_IF;

    IF ipText[tmp_pos - 1] <> 46 THEN
        ipValue := 0;
        RETURN;
    END_IF;

    tmp_pos := tmp_pos + 1;
END_WHILE;

IF tmp_byte_index <> 4 THEN
    ipValue := 0;
    RETURN;
END_IF;

ipValue := (tmp_byte0 * 16777216) OR (tmp_byte1 * 65536) OR (tmp_byte2 * 256) OR tmp_byte3;

END_FUNCTION_BLOCK

(* CONTRACT_RULES [] *)

(* ---- public-medium-08.candidate_02.st ---- *)
FUNCTION_BLOCK IPv4_Parser
VAR_INPUT
    ipText : STRING(254);
END_VAR
VAR_OUTPUT
    ipValue : UDINT;
END_VAR
VAR
    tmp_pos : UDINT;
    tmp_digit : UDINT;
    tmp_val : UDINT;
    tmp_byte0 : UDINT;
    tmp_byte1 : UDINT;
    tmp_byte2 : UDINT;
    tmp_byte3 : UDINT;
    tmp_byte_index : UDINT;
    tmp_text_len : UDINT;
    tmp_char : BYTE;
    tmp_digit_count : UDINT;
END_VAR

(*
ENGINEERING_CONTRACT
PUB001: Four nonempty decimal-digit segments separated by periods
PUB002: Each segment 0-255; invalid/empty → ipValue=0
PUB003: Network byte order: seg1=MSB(31:24), seg4=LSB(7:0)
PUB004: Valid address 0.0.0.0 also produces 0 (boundary case)
*)

tmp_text_len := LEN(ipText);
IF tmp_text_len = 0 OR tmp_text_len > 15 THEN
    ipValue := 0;
    RETURN;
END_IF;

tmp_pos := 1;
tmp_byte_index := 0;

WHILE tmp_byte_index < 4 DO
    tmp_val := 0;
    tmp_digit_count := 0;

    WHILE tmp_pos <= tmp_text_len DO
        tmp_char := ipText[tmp_pos - 1];
        IF tmp_char = 46 THEN
            EXIT;
        END_IF;
        IF tmp_char < 48 OR tmp_char > 57 THEN
            ipValue := 0;
            RETURN;
        END_IF;
        tmp_digit := tmp_char - 48;
        tmp_val := tmp_val * 10 + tmp_digit;
        tmp_digit_count := tmp_digit_count + 1;
        tmp_pos := tmp_pos + 1;
    END_WHILE;

    IF tmp_digit_count = 0 OR tmp_digit_count > 3 THEN
        ipValue := 0;
        RETURN;
    END_IF;

    IF tmp_val > 255 THEN
        ipValue := 0;
        RETURN;
    END_IF;

    IF tmp_byte_index = 0 THEN
        tmp_byte0 := tmp_val;
    ELSIF tmp_byte_index = 1 THEN
        tmp_byte1 := tmp_val;
    ELSIF tmp_byte_index = 2 THEN
        tmp_byte2 := tmp_val;
    ELSIF tmp_byte_index = 3 THEN
        tmp_byte3 := tmp_val;
    END_IF;

    tmp_byte_index := tmp_byte_index + 1;

    IF tmp_pos > tmp_text_len THEN
        EXIT;
    END_IF;

    IF ipText[tmp_pos - 1] <> 46 THEN
        ipValue := 0;
        RETURN;
    END_IF;

    tmp_pos := tmp_pos + 1;
END_WHILE;

IF tmp_byte_index <> 4 THEN
    ipValue := 0;
    RETURN;
END_IF;

ipValue := (tmp_byte0 * 16777216) OR (tmp_byte1 * 65536) OR (tmp_byte2 * 256) OR tmp_byte3;

END_FUNCTION_BLOCK

(* CONTRACT_RULES [] *)

(* ---- public-medium-08.patch_base_02.st ---- *)
FUNCTION_BLOCK IPv4_Parser
VAR_INPUT
    ipText : STRING(254);
END_VAR
VAR_OUTPUT
    ipValue : UDINT;
END_VAR
VAR
    tmp_pos : UDINT;
    tmp_seg : STRING(4);
    tmp_val : UDINT;
    tmp_byte0 : UDINT;
    tmp_byte1 : UDINT;
    tmp_byte2 : UDINT;
    tmp_byte3 : UDINT;
    tmp_byte_index : UDINT;
    tmp_text_len : UDINT;
    tmp_char : BYTE;
    tmp_seg_len : UDINT;
END_VAR

(*
ENGINEERING_CONTRACT
PUB001: Four nonempty decimal-digit segments separated by periods
PUB002: Each segment 0-255; invalid/empty → ipValue=0
PUB003: Network byte order: seg1=MSB(31:24), seg4=LSB(7:0)
PUB004: Valid address 0.0.0.0 also produces 0 (boundary case)
*)

tmp_text_len := LEN(ipText);
IF tmp_text_len = 0 OR tmp_text_len > 15 THEN
    ipValue := 0;
    RETURN;
END_IF;

tmp_pos := 1;
tmp_byte_index := 0;

WHILE tmp_byte_index < 4 DO
    tmp_seg := '';
    tmp_seg_len := 0;

    WHILE tmp_pos <= tmp_text_len DO
        tmp_char := ipText[tmp_pos - 1];
        IF tmp_char = 46 THEN
            EXIT;
        END_IF;
        IF tmp_char < 48 OR tmp_char > 57 THEN
            ipValue := 0;
            RETURN;
        END_IF;
        tmp_seg := CONCAT(tmp_seg, CHR(tmp_char));
        tmp_seg_len := tmp_seg_len + 1;
        tmp_pos := tmp_pos + 1;
    END_WHILE;

    IF tmp_seg_len = 0 OR tmp_seg_len > 3 THEN
        ipValue := 0;
        RETURN;
    END_IF;

    tmp_val := STRING_TO_UDINT(tmp_seg);
    IF tmp_val > 255 THEN
        ipValue := 0;
        RETURN;
    END_IF;

    IF tmp_byte_index = 0 THEN
        tmp_byte0 := tmp_val;
    ELSIF tmp_byte_index = 1 THEN
        tmp_byte1 := tmp_val;
    ELSIF tmp_byte_index = 2 THEN
        tmp_byte2 := tmp_val;
    ELSIF tmp_byte_index = 3 THEN
        tmp_byte3 := tmp_val;
    END_IF;

    tmp_byte_index := tmp_byte_index + 1;

    IF tmp_pos > tmp_text_len THEN
        EXIT;
    END_IF;

    IF ipText[tmp_pos - 1] <> 46 THEN
        ipValue := 0;
        RETURN;
    END_IF;

    tmp_pos := tmp_pos + 1;
END_WHILE;

IF tmp_byte_index <> 4 THEN
    ipValue := 0;
    RETURN;
END_IF;

ipValue := (tmp_byte0 * 16777216) OR (tmp_byte1 * 65536) OR (tmp_byte2 * 256) OR tmp_byte3;

END_FUNCTION_BLOCK

(* CONTRACT_RULES [] *)

(* ---- public-medium-08.patch_base_03.st ---- *)
FUNCTION_BLOCK IPv4_Parser
VAR_INPUT
    ipText : STRING(254);
END_VAR
VAR_OUTPUT
    ipValue : UDINT;
END_VAR
VAR
    tmp_pos : UDINT;
    tmp_digit : UDINT;
    tmp_val : UDINT;
    tmp_byte0 : UDINT;
    tmp_byte1 : UDINT;
    tmp_byte2 : UDINT;
    tmp_byte3 : UDINT;
    tmp_byte_index : UDINT;
    tmp_text_len : UDINT;
    tmp_char : BYTE;
    tmp_digit_count : UDINT;
END_VAR

(*
ENGINEERING_CONTRACT
PUB001: Four nonempty decimal-digit segments separated by periods
PUB002: Each segment 0-255; invalid/empty → ipValue=0
PUB003: Network byte order: seg1=MSB(31:24), seg4=LSB(7:0)
PUB004: Valid address 0.0.0.0 also produces 0 (boundary case)
*)

tmp_text_len := LEN(ipText);
IF tmp_text_len = 0 OR tmp_text_len > 15 THEN
    ipValue := 0;
    RETURN;
END_IF;

tmp_pos := 1;
tmp_byte_index := 0;

WHILE tmp_byte_index < 4 DO
    tmp_val := 0;
    tmp_digit_count := 0;

    WHILE tmp_pos <= tmp_text_len DO
        tmp_char := ipText[tmp_pos - 1];
        IF tmp_char = 46 THEN
            EXIT;
        END_IF;
        IF tmp_char < 48 OR tmp_char > 57 THEN
            ipValue := 0;
            RETURN;
        END_IF;
        tmp_digit := tmp_char - 48;
        tmp_val := tmp_val * 10 + tmp_digit;
        tmp_digit_count := tmp_digit_count + 1;
        tmp_pos := tmp_pos + 1;
    END_WHILE;

    IF tmp_digit_count = 0 OR tmp_digit_count > 3 THEN
        ipValue := 0;
        RETURN;
    END_IF;

    IF tmp_val > 255 THEN
        ipValue := 0;
        RETURN;
    END_IF;

    IF tmp_byte_index = 0 THEN
        tmp_byte0 := tmp_val;
    ELSIF tmp_byte_index = 1 THEN
        tmp_byte1 := tmp_val;
    ELSIF tmp_byte_index = 2 THEN
        tmp_byte2 := tmp_val;
    ELSIF tmp_byte_index = 3 THEN
        tmp_byte3 := tmp_val;
    END_IF;

    tmp_byte_index := tmp_byte_index + 1;

    IF tmp_pos > tmp_text_len THEN
        EXIT;
    END_IF;

    IF ipText[tmp_pos - 1] <> 46 THEN
        ipValue := 0;
        RETURN;
    END_IF;

    tmp_pos := tmp_pos + 1;
END_WHILE;

IF tmp_byte_index <> 4 THEN
    ipValue := 0;
    RETURN;
END_IF;

ipValue := (tmp_byte0 * 16777216) OR (tmp_byte1 * 65536) OR (tmp_byte2 * 256) OR tmp_byte3;

END_FUNCTION_BLOCK

(* CONTRACT_RULES [] *)

(* ---- public-medium-08.patch_base_04.st ---- *)
FUNCTION_BLOCK IPv4_Parser
VAR_INPUT
    ipText : STRING(254);
END_VAR
VAR_OUTPUT
    ipValue : UDINT;
END_VAR
VAR
    tmp_pos : UDINT;
    tmp_digit : UDINT;
    tmp_val : UDINT;
    tmp_byte0 : UDINT;
    tmp_byte1 : UDINT;
    tmp_byte2 : UDINT;
    tmp_byte3 : UDINT;
    tmp_byte_index : UDINT;
    tmp_text_len : UDINT;
    tmp_char : BYTE;
    tmp_digit_count : UDINT;
END_VAR

(*
ENGINEERING_CONTRACT
PUB001: Four nonempty decimal-digit segments separated by periods
PUB002: Each segment 0-255; invalid/empty → ipValue=0
PUB003: Network byte order: seg1=MSB(31:24), seg4=LSB(7:0)
PUB004: Valid address 0.0.0.0 also produces 0 (boundary case)
*)

tmp_text_len := LEN(ipText);
IF tmp_text_len = 0 OR tmp_text_len > 15 THEN
    ipValue := 0;
    RETURN;
END_IF;

tmp_pos := 1;
tmp_byte_index := 0;

WHILE tmp_byte_index < 4 DO
    tmp_val := 0;
    tmp_digit_count := 0;

    WHILE tmp_pos <= tmp_text_len DO
        tmp_char := ipText[tmp_pos - 1];
        IF tmp_char = 46 THEN
            EXIT;
        END_IF;
        IF tmp_char < 48 OR tmp_char > 57 THEN
            ipValue := 0;
            RETURN;
        END_IF;
        tmp_digit := tmp_char - 48;
        tmp_val := tmp_val * 10 + tmp_digit;
        tmp_digit_count := tmp_digit_count + 1;
        tmp_pos := tmp_pos + 1;
    END_WHILE;

    IF tmp_digit_count = 0 OR tmp_digit_count > 3 THEN
        ipValue := 0;
        RETURN;
    END_IF;

    IF tmp_val > 255 THEN
        ipValue := 0;
        RETURN;
    END_IF;

    IF tmp_byte_index = 0 THEN
        tmp_byte0 := tmp_val;
    ELSIF tmp_byte_index = 1 THEN
        tmp_byte1 := tmp_val;
    ELSIF tmp_byte_index = 2 THEN
        tmp_byte2 := tmp_val;
    ELSIF tmp_byte_index = 3 THEN
        tmp_byte3 := tmp_val;
    END_IF;

    tmp_byte_index := tmp_byte_index + 1;

    IF tmp_pos > tmp_text_len THEN
        EXIT;
    END_IF;

    IF ipText[tmp_pos - 1] <> 46 THEN
        ipValue := 0;
        RETURN;
    END_IF;

    tmp_pos := tmp_pos + 1;
END_WHILE;

IF tmp_byte_index <> 4 THEN
    ipValue := 0;
    RETURN;
END_IF;

ipValue := (tmp_byte0 * 16777216) OR (tmp_byte1 * 65536) OR (tmp_byte2 * 256) OR tmp_byte3;

END_FUNCTION_BLOCK

(* CONTRACT_RULES [] *)

(* ---- public-medium-08.raw_candidate_01.st ---- *)
FUNCTION_BLOCK IPv4_Parser
VAR_INPUT
    ipText : STRING(254);
END_VAR
VAR_OUTPUT
    ipValue : UDINT;
END_VAR
VAR
    tmp_pos : UDINT;
    tmp_seg : STRING(4);
    tmp_val : UDINT;
    tmp_byte0 : UDINT;
    tmp_byte1 : UDINT;
    tmp_byte2 : UDINT;
    tmp_byte3 : UDINT;
    tmp_byte_index : UDINT;
    tmp_text_len : UDINT;
    tmp_char : BYTE;
    tmp_seg_len : UDINT;
END_VAR

(*
ENGINEERING_CONTRACT
PUB001: Four nonempty decimal-digit segments separated by periods
PUB002: Each segment 0-255; invalid/empty → ipValue=0
PUB003: Network byte order: seg1=MSB(31:24), seg4=LSB(7:0)
PUB004: Valid address 0.0.0.0 also produces 0 (boundary case)
*)

tmp_text_len := LEN(ipText);
IF tmp_text_len = 0 OR tmp_text_len > 15 THEN
    ipValue := 0;
    RETURN;
END_IF;

tmp_pos := 1;
tmp_byte_index := 0;

WHILE tmp_byte_index < 4 DO
    tmp_seg := '';
    tmp_seg_len := 0;

    WHILE tmp_pos <= tmp_text_len DO
        tmp_char := ipText[tmp_pos - 1];
        IF tmp_char = 46 THEN
            EXIT;
        END_IF
        IF tmp_char < 48 OR tmp_char > 57 THEN
            ipValue := 0;
            RETURN;
        END_IF
        tmp_seg := CONCAT(tmp_seg, CHR(tmp_char));
        tmp_seg_len := tmp_seg_len + 1;
        tmp_pos := tmp_pos + 1;
    END_WHILE

    IF tmp_seg_len = 0 OR tmp_seg_len > 3 THEN
        ipValue := 0;
        RETURN;
    END_IF

    tmp_val := STRING_TO_UDINT(tmp_seg);
    IF tmp_val > 255 THEN
        ipValue := 0;
        RETURN;
    END_IF

    IF tmp_byte_index = 0 THEN
        tmp_byte0 := tmp_val;
    ELSIF tmp_byte_index = 1 THEN
        tmp_byte1 := tmp_val;
    ELSIF tmp_byte_index = 2 THEN
        tmp_byte2 := tmp_val;
    ELSIF tmp_byte_index = 3 THEN
        tmp_byte3 := tmp_val;
    END_IF

    tmp_byte_index := tmp_byte_index + 1;

    IF tmp_pos > tmp_text_len THEN
        EXIT;
    END_IF

    IF ipText[tmp_pos - 1] <> 46 THEN
        ipValue := 0;
        RETURN;
    END_IF

    tmp_pos := tmp_pos + 1;
END_WHILE;

IF tmp_byte_index <> 4 THEN
    ipValue := 0;
    RETURN;
END_IF;

ipValue := (tmp_byte0 * 16777216) OR (tmp_byte1 * 65536) OR (tmp_byte2 * 256) OR tmp_byte3;

END_FUNCTION_BLOCK

(* CONTRACT_RULES [] *)

(* ---- public-medium-08.raw_candidate_02.st ---- *)
FUNCTION_BLOCK IPv4_Parser
VAR_INPUT
    ipText : STRING(254);
END_VAR
VAR_OUTPUT
    ipValue : UDINT;
END_VAR
VAR
    tmp_pos : UDINT;
    tmp_digit : UDINT;
    tmp_val : UDINT;
    tmp_byte0 : UDINT;
    tmp_byte1 : UDINT;
    tmp_byte2 : UDINT;
    tmp_byte3 : UDINT;
    tmp_byte_index : UDINT;
    tmp_text_len : UDINT;
    tmp_char : BYTE;
    tmp_digit_count : UDINT;
END_VAR

(*
ENGINEERING_CONTRACT
PUB001: Four nonempty decimal-digit segments separated by periods
PUB002: Each segment 0-255; invalid/empty → ipValue=0
PUB003: Network byte order: seg1=MSB(31:24), seg4=LSB(7:0)
PUB004: Valid address 0.0.0.0 also produces 0 (boundary case)
*)

tmp_text_len := LEN(ipText);
IF tmp_text_len = 0 OR tmp_text_len > 15 THEN
    ipValue := 0;
    RETURN;
END_IF;

tmp_pos := 1;
tmp_byte_index := 0;

WHILE tmp_byte_index < 4 DO
    tmp_val := 0;
    tmp_digit_count := 0;

    WHILE tmp_pos <= tmp_text_len DO
        tmp_char := ipText[tmp_pos - 1];
        IF tmp_char = 46 THEN
            EXIT;
        END_IF;
        IF tmp_char < 48 OR tmp_char > 57 THEN
            ipValue := 0;
            RETURN;
        END_IF;
        tmp_digit := tmp_char - 48;
        tmp_val := tmp_val * 10 + tmp_digit;
        tmp_digit_count := tmp_digit_count + 1;
        tmp_pos := tmp_pos + 1;
    END_WHILE;

    IF tmp_digit_count = 0 OR tmp_digit_count > 3 THEN
        ipValue := 0;
        RETURN;
    END_IF;

    IF tmp_val > 255 THEN
        ipValue := 0;
        RETURN;
    END_IF;

    IF tmp_byte_index = 0 THEN
        tmp_byte0 := tmp_val;
    ELSIF tmp_byte_index = 1 THEN
        tmp_byte1 := tmp_val;
    ELSIF tmp_byte_index = 2 THEN
        tmp_byte2 := tmp_val;
    ELSIF tmp_byte_index = 3 THEN
        tmp_byte3 := tmp_val;
    END_IF;

    tmp_byte_index := tmp_byte_index + 1;

    IF tmp_pos > tmp_text_len THEN
        EXIT;
    END_IF;

    IF ipText[tmp_pos - 1] <> 46 THEN
        ipValue := 0;
        RETURN;
    END_IF;

    tmp_pos := tmp_pos + 1;
END_WHILE;

IF tmp_byte_index <> 4 THEN
    ipValue := 0;
    RETURN;
END_IF;

ipValue := (tmp_byte0 * 16777216) OR (tmp_byte1 * 65536) OR (tmp_byte2 * 256) OR tmp_byte3;

END_FUNCTION_BLOCK

(* CONTRACT_RULES [] *)

(* ---- self-easy-01.candidate_01.st ---- *)
(* ENGINEERING_CONTRACT
================================================================
| Output/State    | Activation           | Retention          | Reset/Deactivation       | Priority | Units          |
|-----------------|----------------------|--------------------|--------------------------|----------|----------------|
| avgOut          | enable AND count>0   | prev value         | enable=FALSE OR count=0  | Same-scan| REAL           |
|                 | AND avgEnable=TRUE   |                    | OR avgEnable=FALSE       |          |                |
================================================================
Behavior:
- avgOut updates only when: enable=TRUE, count>0, avgEnable=TRUE
- avgOut holds (retention) when: enable=FALSE, OR count<=0, OR avgEnable=FALSE
- Sum uses DINT to prevent overflow; division by clipped count (max 8, min 1)
- No NaN possible: division only when count >= 1

*)

(* CONTRACT_RULES [] *)

FUNCTION_BLOCK FB
VAR
    tmp_sum : DINT := 0;
    tmp_i   : INT  := 0;
END_VAR
VAR_INPUT
    enable     : BOOL;
    values     : ARRAY[1..8] OF INT;
    count      : INT;
    avgEnable  : BOOL;
END_VAR
VAR_OUTPUT
    avgOut : REAL := 0.0;
END_VAR

IF enable AND avgEnable AND count > 0 THEN
    tmp_sum := 0;
    FOR tmp_i := 1 TO MIN(count, 8) DO
        tmp_sum := tmp_sum + INT_TO_DINT(values[tmp_i]);
    END_FOR;
    avgOut := DINT_TO_REAL(tmp_sum) / INT_TO_REAL(MAX(count, 1));
END_IF;
END_FUNCTION_BLOCK

(* ---- self-easy-01.patch_base_02.st ---- *)
(* ENGINEERING_CONTRACT
================================================================
| Output/State    | Activation           | Retention          | Reset/Deactivation       | Priority | Units          |
|-----------------|----------------------|--------------------|--------------------------|----------|----------------|
| avgOut          | enable AND count>0   | prev value         | enable=FALSE OR count=0  | Same-scan| REAL           |
|                 | AND avgEnable=TRUE   |                    | OR avgEnable=FALSE       |          |                |
================================================================
Behavior:
- avgOut updates only when: enable=TRUE, count>0, avgEnable=TRUE
- avgOut holds (retention) when: enable=FALSE, OR count<=0, OR avgEnable=FALSE
- Sum uses DINT to prevent overflow; division by clipped count (max 8, min 1)
- No NaN possible: division only when count >= 1

*)

(* CONTRACT_RULES [] *)

FUNCTION_BLOCK FB
VAR
    tmp_sum : DINT := 0;
    tmp_i   : INT  := 0;
END_VAR
VAR_INPUT
    enable     : BOOL;
    values     : ARRAY[1..8] OF INT;
    count      : INT;
    avgEnable  : BOOL;
END_VAR
VAR_OUTPUT
    avgOut : REAL := 0.0;
END_VAR

IF enable AND avgEnable AND count > 0 THEN
    tmp_sum := 0;
    FOR tmp_i := 1 TO MIN(count, 8) DO
        tmp_sum := tmp_sum + INT_TO_DINT(values[tmp_i]);
    END_FOR;
    avgOut := DINT_TO_REAL(tmp_sum) / INT_TO_REAL(MAX(count, 1));
END_IF;
END_FUNCTION_BLOCK

(* ---- self-easy-01.patch_base_03.st ---- *)
(* ENGINEERING_CONTRACT
================================================================
| Output/State    | Activation           | Retention          | Reset/Deactivation       | Priority | Units          |
|-----------------|----------------------|--------------------|--------------------------|----------|----------------|
| avgOut          | enable AND count>0   | prev value         | enable=FALSE OR count=0  | Same-scan| REAL           |
|                 | AND avgEnable=TRUE   |                    | OR avgEnable=FALSE       |          |                |
================================================================
Behavior:
- avgOut updates only when: enable=TRUE, count>0, avgEnable=TRUE
- avgOut holds (retention) when: enable=FALSE, OR count<=0, OR avgEnable=FALSE
- Sum uses DINT to prevent overflow; division by clipped count (max 8, min 1)
- No NaN possible: division only when count >= 1

*)

(* CONTRACT_RULES [] *)

FUNCTION_BLOCK FB
VAR
    tmp_sum : DINT := 0;
    tmp_i   : INT  := 0;
END_VAR
VAR_INPUT
    enable     : BOOL;
    values     : ARRAY[1..8] OF INT;
    count      : INT;
    avgEnable  : BOOL;
END_VAR
VAR_OUTPUT
    avgOut : REAL := 0.0;
END_VAR

IF enable AND avgEnable AND count > 0 THEN
    tmp_sum := 0;
    FOR tmp_i := 1 TO MIN(count, 8) DO
        tmp_sum := tmp_sum + INT_TO_DINT(values[tmp_i]);
    END_FOR;
    avgOut := DINT_TO_REAL(tmp_sum) / INT_TO_REAL(MAX(count, 1));
END_IF;
END_FUNCTION_BLOCK

(* ---- self-easy-01.raw_candidate_01.st ---- *)
(* ENGINEERING_CONTRACT
================================================================
| Output/State    | Activation           | Retention          | Reset/Deactivation       | Priority | Units          |
|-----------------|----------------------|--------------------|--------------------------|----------|----------------|
| avgOut          | enable AND count>0   | prev value         | enable=FALSE OR count=0  | Same-scan| REAL           |
|                 | AND avgEnable=TRUE   |                    | OR avgEnable=FALSE       |          |                |
================================================================
Behavior:
- avgOut updates only when: enable=TRUE, count>0, avgEnable=TRUE
- avgOut holds (retention) when: enable=FALSE, OR count<=0, OR avgEnable=FALSE
- Sum uses DINT to prevent overflow; division by clipped count (max 8, min 1)
- No NaN possible: division only when count >= 1

*)

(* CONTRACT_RULES [] *)

FUNCTION_BLOCK FB
VAR
    tmp_sum : DINT := 0;
    tmp_i   : INT  := 0;
END_VAR
VAR_INPUT
    enable     : BOOL;
    values     : ARRAY[1..8] OF INT;
    count      : INT;
    avgEnable  : BOOL;
END_VAR
VAR_OUTPUT
    avgOut : REAL := 0.0;
END_VAR

IF enable AND avgEnable AND count > 0 THEN
    tmp_sum := 0;
    FOR tmp_i := 1 TO MIN(count, 8) DO
        tmp_sum := tmp_sum + INT_TO_DINT(values[tmp_i]);
    END_FOR;
    avgOut := DINT_TO_REAL(tmp_sum) / INT_TO_REAL(MAX(count, 1));
END_IF;
END_FUNCTION_BLOCK

(* ---- self-easy-02.candidate_01.st ---- *)
FUNCTION_BLOCK FB
VAR_INPUT
    tankLevel   : REAL;
    outletFlow  : REAL;
    inletPermit : BOOL;
    resetBtn    : BOOL;
END_VAR
VAR_OUTPUT
    pumpRun         : BOOL;
    alarmHigh       : BOOL;
    alarmLow        : BOOL;
    outletValveOpen : BOOL;
END_VAR
VAR
    prevResetBtn : BOOL := FALSE;
    tmpRising    : BOOL;
END_VAR

(*
ENGINEERING_CONTRACT
============================================================
Output | Activation         | Retention        | Reset/Deactivation    | Same-scan Priority | Units
-------|--------------------|------------------|-----------------------|--------------------|-------------
alarmHigh | tankLevel>=85.0   | hold until reset | rising(resetBtn) & tankLevel<85.0 | danger prioritizes over reset | BOOL latch
alarmLow  | tankLevel<=15.0   | hold until reset | rising(resetBtn) & tankLevel>15.0 | danger prioritizes over reset | BOOL latch
pumpRun   | inletPermit & !alarmHigh & !alarmLow | no retention | deasserts when alarm set | alarm blocks pump | combinational
outletValveOpen | !alarmLow    | no retention    | asserts when alarmLow=FALSE | alarmLow→closed | combinational inverse
============================================================
PUB: alarmHigh set by PUB001, alarmLow set by PUB003
PUB: alarmHigh reset by PUB005 (rising edge check), alarmLow reset by PUB005
PUB: pumpRun = inletPermit AND no alarms (PUB003, PUB007, PUB019, PUB026)
PUB: outletValveOpen = NOT alarmLow (PUB004, PUB027)
============================================================
*)

(* CONTRACT_RULES [] *)

tmpRising := resetBtn AND NOT prevResetBtn;

alarmHigh := alarmHigh OR (tankLevel >= 85.0);
IF tmpRising THEN
    IF tankLevel < 85.0 THEN
        alarmHigh := FALSE;
    END_IF;
END_IF;

alarmLow := alarmLow OR (tankLevel <= 15.0);
IF tmpRising THEN
    IF tankLevel > 15.0 THEN
        alarmLow := FALSE;
    END_IF;
END_IF;

prevResetBtn := resetBtn;

pumpRun := inletPermit AND NOT alarmHigh AND NOT alarmLow;

outletValveOpen := NOT alarmLow;

END_FUNCTION_BLOCK

(* ---- self-easy-02.raw_candidate_01.st ---- *)
FUNCTION_BLOCK FB
VAR_INPUT
    tankLevel   : REAL;
    outletFlow  : REAL;
    inletPermit : BOOL;
    resetBtn    : BOOL;
END_VAR
VAR_OUTPUT
    pumpRun         : BOOL;
    alarmHigh       : BOOL;
    alarmLow        : BOOL;
    outletValveOpen : BOOL;
END_VAR
VAR
    prevResetBtn : BOOL := FALSE;
    tmpRising    : BOOL;
END_VAR

(*
ENGINEERING_CONTRACT
============================================================
Output | Activation         | Retention        | Reset/Deactivation    | Same-scan Priority | Units
-------|--------------------|------------------|-----------------------|--------------------|-------------
alarmHigh | tankLevel>=85.0   | hold until reset | rising(resetBtn) & tankLevel<85.0 | danger prioritizes over reset | BOOL latch
alarmLow  | tankLevel<=15.0   | hold until reset | rising(resetBtn) & tankLevel>15.0 | danger prioritizes over reset | BOOL latch
pumpRun   | inletPermit & !alarmHigh & !alarmLow | no retention | deasserts when alarm set | alarm blocks pump | combinational
outletValveOpen | !alarmLow    | no retention    | asserts when alarmLow=FALSE | alarmLow→closed | combinational inverse
============================================================
PUB: alarmHigh set by PUB001, alarmLow set by PUB003
PUB: alarmHigh reset by PUB005 (rising edge check), alarmLow reset by PUB005
PUB: pumpRun = inletPermit AND no alarms (PUB003, PUB007, PUB019, PUB026)
PUB: outletValveOpen = NOT alarmLow (PUB004, PUB027)
============================================================
*)

(* CONTRACT_RULES [] *)

tmpRising := resetBtn AND NOT prevResetBtn;

alarmHigh := alarmHigh OR (tankLevel >= 85.0);
IF tmpRising THEN
    IF tankLevel < 85.0 THEN
        alarmHigh := FALSE;
    END_IF;
END_IF;

alarmLow := alarmLow OR (tankLevel <= 15.0);
IF tmpRising THEN
    IF tankLevel > 15.0 THEN
        alarmLow := FALSE;
    END_IF;
END_IF;

prevResetBtn := resetBtn;

pumpRun := inletPermit AND NOT alarmHigh AND NOT alarmLow;

outletValveOpen := NOT alarmLow;

END_FUNCTION_BLOCK

(* ---- self-hard-01.candidate_01.st ---- *)
(* ENGINEERING_CONTRACT
 * alarmActive: activation=flowLow rising edge(PUB001), retention=until ack when cleared, reset=ackBtn rising when active & !flowLow(PUB010)
 * alarmAcked: activation=condition cleared after active(PUB002-003), retention=until alarmActive clears, reset=same-scan with alarmActive(PUB010)
 * highHigh: activation=!sensorOK(PUB004), retention=while !sensorOK, reset=sensorOK recovery(PUB005)
 * Units: BOOL states, edge-detect via local prev variables, no timers
 *)
(* CONTRACT_RULES [{"kind":"hold_until_reset","output":"alarmActive","set_input":"flowLow","reset_input":"ackBtn"},{"kind":"hold_until_reset","output":"alarmAcked","set_input":"flowLow","reset_input":"ackBtn"}] *)

FUNCTION_BLOCK FB
VAR_INPUT
    flowLow   : BOOL;
    ackBtn    : BOOL;
    sensorOK  : BOOL;
END_VAR
VAR_OUTPUT
    alarmActive : BOOL;
    alarmAcked  : BOOL;
    highHigh    : BOOL;
END_VAR
VAR
    prev_ackBtn   : BOOL;
    prev_flowLow  : BOOL;
END_VAR

    IF ackBtn AND NOT prev_ackBtn THEN
        IF alarmActive THEN
            IF flowLow THEN
                alarmAcked := TRUE;
            ELSE
                alarmActive := FALSE;
                alarmAcked  := FALSE;
            END_IF;
        END_IF;
    ELSIF flowLow AND NOT prev_flowLow THEN
        alarmActive := TRUE;
        alarmAcked  := FALSE;
    ELSIF NOT flowLow AND alarmActive AND alarmAcked THEN
        alarmActive := FALSE;
        alarmAcked  := FALSE;
    END_IF;

    highHigh := NOT sensorOK;

    prev_ackBtn  := ackBtn;
    prev_flowLow := flowLow;
END_FUNCTION_BLOCK

(* ---- self-hard-01.patch_base_02.st ---- *)
(* ENGINEERING_CONTRACT
 * alarmActive: activation=flowLow rising edge(PUB001), retention=until ack when cleared, reset=ackBtn rising when active & !flowLow(PUB010)
 * alarmAcked: activation=condition cleared after active(PUB002-003), retention=until alarmActive clears, reset=same-scan with alarmActive(PUB010)
 * highHigh: activation=!sensorOK(PUB004), retention=while !sensorOK, reset=sensorOK recovery(PUB005)
 * Units: BOOL states, edge-detect via local prev variables, no timers
 *)
(* CONTRACT_RULES [{"kind":"hold_until_reset","output":"alarmActive","set_input":"flowLow","reset_input":"ackBtn"},{"kind":"hold_until_reset","output":"alarmAcked","set_input":"flowLow","reset_input":"ackBtn"}] *)

FUNCTION_BLOCK FB
VAR_INPUT
    flowLow   : BOOL;
    ackBtn    : BOOL;
    sensorOK  : BOOL;
END_VAR
VAR_OUTPUT
    alarmActive : BOOL;
    alarmAcked  : BOOL;
    highHigh    : BOOL;
END_VAR
VAR
    prev_ackBtn   : BOOL;
    prev_flowLow  : BOOL;
END_VAR

    IF ackBtn AND NOT prev_ackBtn THEN
        IF alarmActive THEN
            IF flowLow THEN
                alarmAcked := TRUE;
            ELSE
                alarmActive := FALSE;
                alarmAcked  := FALSE;
            END_IF;
        END_IF;
    ELSIF flowLow AND NOT prev_flowLow THEN
        alarmActive := TRUE;
        alarmAcked  := FALSE;
    ELSIF NOT flowLow AND alarmActive AND alarmAcked THEN
        alarmActive := FALSE;
        alarmAcked  := FALSE;
    END_IF;

    highHigh := NOT sensorOK;

    prev_ackBtn  := ackBtn;
    prev_flowLow := flowLow;
END_FUNCTION_BLOCK

(* ---- self-hard-01.patch_base_03.st ---- *)
(* ENGINEERING_CONTRACT
 * alarmActive: activation=flowLow rising edge(PUB001), retention=until ack when cleared, reset=ackBtn rising when active & !flowLow(PUB010)
 * alarmAcked: activation=condition cleared after active(PUB002-003), retention=until alarmActive clears, reset=same-scan with alarmActive(PUB010)
 * highHigh: activation=!sensorOK(PUB004), retention=while !sensorOK, reset=sensorOK recovery(PUB005)
 * Units: BOOL states, edge-detect via local prev variables, no timers
 *)
(* CONTRACT_RULES [{"kind":"hold_until_reset","output":"alarmActive","set_input":"flowLow","reset_input":"ackBtn"},{"kind":"hold_until_reset","output":"alarmAcked","set_input":"flowLow","reset_input":"ackBtn"}] *)

FUNCTION_BLOCK FB
VAR_INPUT
    flowLow   : BOOL;
    ackBtn    : BOOL;
    sensorOK  : BOOL;
END_VAR
VAR_OUTPUT
    alarmActive : BOOL;
    alarmAcked  : BOOL;
    highHigh    : BOOL;
END_VAR
VAR
    prev_ackBtn   : BOOL;
    prev_flowLow  : BOOL;
END_VAR

    IF ackBtn AND NOT prev_ackBtn THEN
        IF alarmActive THEN
            IF flowLow THEN
                alarmAcked := TRUE;
            ELSE
                alarmActive := FALSE;
                alarmAcked  := FALSE;
            END_IF;
        END_IF;
    ELSIF flowLow AND NOT prev_flowLow THEN
        alarmActive := TRUE;
        alarmAcked  := FALSE;
    ELSIF NOT flowLow AND alarmActive AND alarmAcked THEN
        alarmActive := FALSE;
        alarmAcked  := FALSE;
    END_IF;

    highHigh := NOT sensorOK;

    prev_ackBtn  := ackBtn;
    prev_flowLow := flowLow;
END_FUNCTION_BLOCK

(* ---- self-hard-01.raw_candidate_01.st ---- *)
(* ENGINEERING_CONTRACT
 * alarmActive: activation=flowLow rising edge(PUB001), retention=until ack when cleared, reset=ackBtn rising when active & !flowLow(PUB010)
 * alarmAcked: activation=condition cleared after active(PUB002-003), retention=until alarmActive clears, reset=same-scan with alarmActive(PUB010)
 * highHigh: activation=!sensorOK(PUB004), retention=while !sensorOK, reset=sensorOK recovery(PUB005)
 * Units: BOOL states, edge-detect via local prev variables, no timers
 *)
(* CONTRACT_RULES [{"kind":"hold_until_reset","output":"alarmActive","set_input":"flowLow","reset_input":"ackBtn"},{"kind":"hold_until_reset","output":"alarmAcked","set_input":"flowLow","reset_input":"ackBtn"}] *)

FUNCTION_BLOCK FB
VAR_INPUT
    flowLow   : BOOL;
    ackBtn    : BOOL;
    sensorOK  : BOOL;
END_VAR
VAR_OUTPUT
    alarmActive : BOOL;
    alarmAcked  : BOOL;
    highHigh    : BOOL;
END_VAR
VAR
    prev_ackBtn   : BOOL;
    prev_flowLow  : BOOL;
END_VAR

    IF ackBtn AND NOT prev_ackBtn THEN
        IF alarmActive THEN
            IF flowLow THEN
                alarmAcked := TRUE;
            ELSE
                alarmActive := FALSE;
                alarmAcked  := FALSE;
            END_IF;
        END_IF;
    ELSIF flowLow AND NOT prev_flowLow THEN
        alarmActive := TRUE;
        alarmAcked  := FALSE;
    ELSIF NOT flowLow AND alarmActive AND alarmAcked THEN
        alarmActive := FALSE;
        alarmAcked  := FALSE;
    END_IF;

    highHigh := NOT sensorOK;

    prev_ackBtn  := ackBtn;
    prev_flowLow := flowLow;
END_FUNCTION_BLOCK

(* ---- self-hard-02.candidate_01.st ---- *)
(* ENGINEERING_CONTRACT:
 * Phase activation:
 *   - Phase 0 (IDLE): Initial and idle; no counting, waiting for start
 *   - Phase 1 (HEATING): Active; elapsed increments, transitions to phase 2 on pv>=setpoint
 *   - Phase 2 (HOLDING): Active; elapsed increments, retained until timeout/abort/start
 *   - Phase 3 (COMPLETE): Retention; elapsed/timeout frozen until new start or abort
 *   - Phase 9 (ABORTED): Retention; elapsed/timeout frozen until new start
 *
 * Priority per scan (same-scan order):
 *   1. abortBtn=TRUE  → phase=9, preserve elapsed/timeout
 *   2. startBtn rising edge (no abort) → phase=1, elapsed=0, timeout=FALSE
 *   3. running (no abort, no start edge) → count if prev phase 1/2, else hold
 *
 * Counting:
 *   - Start scan: elapsed=0 (not counted)
 *   - Running scans: elapsed += 1 while prev phase 1 or 2
 *   - maxDuration: positive INT, comparison elapsed >= maxDuration triggers timeout
 *
 * Units: maxDuration in scan cycles, elapsed in scan cycles
 * Reset: Only new start rising edge (with no abort) clears elapsed/timeout
 *)

FUNCTION_BLOCK FB
VAR_INPUT
    startBtn    : BOOL;
    abortBtn    : BOOL;
    setpoint    : REAL;
    pv          : REAL;
    maxDuration : INT;
END_VAR

VAR_OUTPUT
    elapsed : INT := 0;
    phase   : INT := 0;
    timeout : BOOL := FALSE;
END_VAR

VAR
    prev_startBtn : BOOL := FALSE;
END_VAR

VAR
    startRising : BOOL;
    prev_phase  : INT;
END_VAR

// Detect rising edge of startBtn for this scan
startRising := startBtn AND NOT prev_startBtn;
prev_phase  := phase;

// Priority 1: Abort (highest)
IF abortBtn THEN
    phase := 9;
    // elapsed and timeout are preserved
    prev_startBtn := startBtn;
    RETURN;
END_IF;

// Priority 2: New start rising edge (no abort)
IF startRising THEN
    phase   := 1;
    elapsed := 0;
    timeout := FALSE;
    prev_startBtn := startBtn;
    RETURN;
END_IF;

// Priority 3: Running / frozen states (no abort, no new start edge)
IF prev_phase = 1 OR prev_phase = 2 THEN
    // Running: increment elapsed
    elapsed := elapsed + 1;

    IF elapsed >= maxDuration THEN
        // Timeout: enter complete state
        timeout := TRUE;
        phase   := 3;
    ELSE
        // Not yet timed out: determine phase
        IF pv >= setpoint THEN
            phase := 2;          // pv达标，保持保温
        ELSE
            phase := 1;          // 仍处于升温
        END_IF;
    END_IF;
ELSE
    // Frozen: idle (phase=0), complete (phase=3), or aborted (phase=9)
    // phase and timeout retain their values
END_IF;

prev_startBtn := startBtn;

END_FUNCTION_BLOCK

(* ---- self-hard-02.candidate_03.st ---- *)
(* ENGINEERING_CONTRACT:
 * Phase activation:
 *   - Phase 0 (IDLE): Initial and idle; no counting, waiting for start
 *   - Phase 1 (HEATING): Active; elapsed increments, transitions to phase 2 on pv>=setpoint
 *   - Phase 2 (HOLDING): Active; elapsed increments, retained until timeout/abort/start
 *   - Phase 3 (COMPLETE): Retention; elapsed/timeout frozen until new start or abort
 *   - Phase 9 (ABORTED): Retention; elapsed/timeout frozen until new start
 *
 * Priority per scan (same-scan order):
 *   1. abortBtn=TRUE  → phase=9, preserve elapsed/timeout
 *   2. startBtn rising edge (no abort) → phase=1, elapsed=0, timeout=FALSE
 *   3. running (no abort, no start edge) → count if prev phase 1/2, else hold
 *
 * Counting:
 *   - Start scan: elapsed=0 (not counted)
 *   - Running scans: elapsed += 1 while prev phase 1 or 2
 *   - maxDuration: positive INT, comparison elapsed >= maxDuration triggers timeout
 *
 * Units: maxDuration in scan cycles, elapsed in scan cycles
 * Reset: Only new start rising edge (with no abort) clears elapsed/timeout
 *)

FUNCTION_BLOCK FB
VAR_INPUT
    startBtn    : BOOL;
    abortBtn    : BOOL;
    setpoint    : REAL;
    pv          : REAL;
    maxDuration : INT;
END_VAR

VAR_OUTPUT
    elapsed : INT := 0;
    phase   : INT := 0;
    timeout : BOOL := FALSE;
END_VAR

VAR
    prev_startBtn : BOOL := FALSE;
    startRising   : BOOL;
    prev_phase    : INT;
END_VAR

// Detect rising edge of startBtn for this scan
startRising := startBtn AND NOT prev_startBtn;
prev_phase  := phase;

// Priority 1: Abort (highest)
IF abortBtn THEN
    phase := 9;
    prev_startBtn := startBtn;
    RETURN;
END_IF;

// Priority 2: New start rising edge (no abort)
IF startRising THEN
    phase   := 1;
    elapsed := 0;
    timeout := FALSE;
    prev_startBtn := startBtn;
    RETURN;
END_IF;

// Priority 3: Running / frozen states (no abort, no new start edge)
IF prev_phase = 1 OR prev_phase = 2 THEN
    // Running: increment elapsed
    elapsed := elapsed + 1;

    IF elapsed >= maxDuration THEN
        // Timeout: enter complete state
        timeout := TRUE;
        phase   := 3;
    ELSE
        // Not yet timed out: determine phase
        IF pv >= setpoint THEN
            phase := 2;
        ELSE
            phase := 1;
        END_IF;
    END_IF;
END_IF;

prev_startBtn := startBtn;

END_FUNCTION_BLOCK

(* ---- self-hard-02.patch_base_02.st ---- *)
(* ENGINEERING_CONTRACT:
 * Phase activation:
 *   - Phase 0 (IDLE): Initial and idle; no counting, waiting for start
 *   - Phase 1 (HEATING): Active; elapsed increments, transitions to phase 2 on pv>=setpoint
 *   - Phase 2 (HOLDING): Active; elapsed increments, retained until timeout/abort/start
 *   - Phase 3 (COMPLETE): Retention; elapsed/timeout frozen until new start or abort
 *   - Phase 9 (ABORTED): Retention; elapsed/timeout frozen until new start
 *
 * Priority per scan (same-scan order):
 *   1. abortBtn=TRUE  → phase=9, preserve elapsed/timeout
 *   2. startBtn rising edge (no abort) → phase=1, elapsed=0, timeout=FALSE
 *   3. running (no abort, no start edge) → count if prev phase 1/2, else hold
 *
 * Counting:
 *   - Start scan: elapsed=0 (not counted)
 *   - Running scans: elapsed += 1 while prev phase 1 or 2
 *   - maxDuration: positive INT, comparison elapsed >= maxDuration triggers timeout
 *
 * Units: maxDuration in scan cycles, elapsed in scan cycles
 * Reset: Only new start rising edge (with no abort) clears elapsed/timeout
 *)

FUNCTION_BLOCK FB
VAR_INPUT
    startBtn    : BOOL;
    abortBtn    : BOOL;
    setpoint    : REAL;
    pv          : REAL;
    maxDuration : INT;
END_VAR

VAR_OUTPUT
    elapsed : INT := 0;
    phase   : INT := 0;
    timeout : BOOL := FALSE;
END_VAR

VAR
    prev_startBtn : BOOL := FALSE;
END_VAR

VAR
    startRising : BOOL;
    prev_phase  : INT;
END_VAR

// Detect rising edge of startBtn for this scan
startRising := startBtn AND NOT prev_startBtn;
prev_phase  := phase;

// Priority 1: Abort (highest)
IF abortBtn THEN
    phase := 9;
    // elapsed and timeout are preserved
    prev_startBtn := startBtn;
    RETURN;
END_IF;

// Priority 2: New start rising edge (no abort)
IF startRising THEN
    phase   := 1;
    elapsed := 0;
    timeout := FALSE;
    prev_startBtn := startBtn;
    RETURN;
END_IF;

// Priority 3: Running / frozen states (no abort, no new start edge)
IF prev_phase = 1 OR prev_phase = 2 THEN
    // Running: increment elapsed
    elapsed := elapsed + 1;

    IF elapsed >= maxDuration THEN
        // Timeout: enter complete state
        timeout := TRUE;
        phase   := 3;
    ELSE
        // Not yet timed out: determine phase
        IF pv >= setpoint THEN
            phase := 2;          // pv达标，保持保温
        ELSE
            phase := 1;          // 仍处于升温
        END_IF;
    END_IF;
ELSE
    // Frozen: idle (phase=0), complete (phase=3), or aborted (phase=9)
    // phase and timeout retain their values
END_IF;

prev_startBtn := startBtn;

END_FUNCTION_BLOCK

(* ---- self-hard-02.patch_base_03.st ---- *)
(* ENGINEERING_CONTRACT:
 * Phase activation:
 *   - Phase 0 (IDLE): Initial and idle; no counting, waiting for start
 *   - Phase 1 (HEATING): Active; elapsed increments, transitions to phase 2 on pv>=setpoint
 *   - Phase 2 (HOLDING): Active; elapsed increments, retained until timeout/abort/start
 *   - Phase 3 (COMPLETE): Retention; elapsed/timeout frozen until new start or abort
 *   - Phase 9 (ABORTED): Retention; elapsed/timeout frozen until new start
 *
 * Priority per scan (same-scan order):
 *   1. abortBtn=TRUE  → phase=9, preserve elapsed/timeout
 *   2. startBtn rising edge (no abort) → phase=1, elapsed=0, timeout=FALSE
 *   3. running (no abort, no start edge) → count if prev phase 1/2, else hold
 *
 * Counting:
 *   - Start scan: elapsed=0 (not counted)
 *   - Running scans: elapsed += 1 while prev phase 1 or 2
 *   - maxDuration: positive INT, comparison elapsed >= maxDuration triggers timeout
 *
 * Units: maxDuration in scan cycles, elapsed in scan cycles
 * Reset: Only new start rising edge (with no abort) clears elapsed/timeout
 *)

FUNCTION_BLOCK FB
VAR_INPUT
    startBtn    : BOOL;
    abortBtn    : BOOL;
    setpoint    : REAL;
    pv          : REAL;
    maxDuration : INT;
END_VAR

VAR_OUTPUT
    elapsed : INT := 0;
    phase   : INT := 0;
    timeout : BOOL := FALSE;
END_VAR

VAR
    prev_startBtn : BOOL := FALSE;
END_VAR

VAR
    startRising : BOOL;
    prev_phase  : INT;
END_VAR

// Detect rising edge of startBtn for this scan
startRising := startBtn AND NOT prev_startBtn;
prev_phase  := phase;

// Priority 1: Abort (highest)
IF abortBtn THEN
    phase := 9;
    // elapsed and timeout are preserved
    prev_startBtn := startBtn;
    RETURN;
END_IF;

// Priority 2: New start rising edge (no abort)
IF startRising THEN
    phase   := 1;
    elapsed := 0;
    timeout := FALSE;
    prev_startBtn := startBtn;
    RETURN;
END_IF;

// Priority 3: Running / frozen states (no abort, no new start edge)
IF prev_phase = 1 OR prev_phase = 2 THEN
    // Running: increment elapsed
    elapsed := elapsed + 1;

    IF elapsed >= maxDuration THEN
        // Timeout: enter complete state
        timeout := TRUE;
        phase   := 3;
    ELSE
        // Not yet timed out: determine phase
        IF pv >= setpoint THEN
            phase := 2;          // pv达标，保持保温
        ELSE
            phase := 1;          // 仍处于升温
        END_IF;
    END_IF;
ELSE
    // Frozen: idle (phase=0), complete (phase=3), or aborted (phase=9)
    // phase and timeout retain their values
END_IF;

prev_startBtn := startBtn;

END_FUNCTION_BLOCK

(* ---- self-hard-02.patch_base_04.st ---- *)
(* ENGINEERING_CONTRACT:
 * Phase activation:
 *   - Phase 0 (IDLE): Initial and idle; no counting, waiting for start
 *   - Phase 1 (HEATING): Active; elapsed increments, transitions to phase 2 on pv>=setpoint
 *   - Phase 2 (HOLDING): Active; elapsed increments, retained until timeout/abort/start
 *   - Phase 3 (COMPLETE): Retention; elapsed/timeout frozen until new start or abort
 *   - Phase 9 (ABORTED): Retention; elapsed/timeout frozen until new start
 *
 * Priority per scan (same-scan order):
 *   1. abortBtn=TRUE  → phase=9, preserve elapsed/timeout
 *   2. startBtn rising edge (no abort) → phase=1, elapsed=0, timeout=FALSE
 *   3. running (no abort, no start edge) → count if prev phase 1/2, else hold
 *
 * Counting:
 *   - Start scan: elapsed=0 (not counted)
 *   - Running scans: elapsed += 1 while prev phase 1 or 2
 *   - maxDuration: positive INT, comparison elapsed >= maxDuration triggers timeout
 *
 * Units: maxDuration in scan cycles, elapsed in scan cycles
 * Reset: Only new start rising edge (with no abort) clears elapsed/timeout
 *)

FUNCTION_BLOCK FB
VAR_INPUT
    startBtn    : BOOL;
    abortBtn    : BOOL;
    setpoint    : REAL;
    pv          : REAL;
    maxDuration : INT;
END_VAR

VAR_OUTPUT
    elapsed : INT := 0;
    phase   : INT := 0;
    timeout : BOOL := FALSE;
END_VAR

VAR
    prev_startBtn : BOOL := FALSE;
    startRising   : BOOL;
    prev_phase    : INT;
END_VAR

// Detect rising edge of startBtn for this scan
startRising := startBtn AND NOT prev_startBtn;
prev_phase  := phase;

// Priority 1: Abort (highest)
IF abortBtn THEN
    phase := 9;
    prev_startBtn := startBtn;
    RETURN;
END_IF;

// Priority 2: New start rising edge (no abort)
IF startRising THEN
    phase   := 1;
    elapsed := 0;
    timeout := FALSE;
    prev_startBtn := startBtn;
    RETURN;
END_IF;

// Priority 3: Running / frozen states (no abort, no new start edge)
IF prev_phase = 1 OR prev_phase = 2 THEN
    // Running: increment elapsed
    elapsed := elapsed + 1;

    IF elapsed >= maxDuration THEN
        // Timeout: enter complete state
        timeout := TRUE;
        phase   := 3;
    ELSE
        // Not yet timed out: determine phase
        IF pv >= setpoint THEN
            phase := 2;
        ELSE
            phase := 1;
        END_IF;
    END_IF;
END_IF;

prev_startBtn := startBtn;

END_FUNCTION_BLOCK

(* ---- self-hard-02.raw_candidate_01.st ---- *)
(* ENGINEERING_CONTRACT:
 * Phase activation:
 *   - Phase 0 (IDLE): Initial and idle; no counting, waiting for start
 *   - Phase 1 (HEATING): Active; elapsed increments, transitions to phase 2 on pv>=setpoint
 *   - Phase 2 (HOLDING): Active; elapsed increments, retained until timeout/abort/start
 *   - Phase 3 (COMPLETE): Retention; elapsed/timeout frozen until new start or abort
 *   - Phase 9 (ABORTED): Retention; elapsed/timeout frozen until new start
 *
 * Priority per scan (same-scan order):
 *   1. abortBtn=TRUE  → phase=9, preserve elapsed/timeout
 *   2. startBtn rising edge (no abort) → phase=1, elapsed=0, timeout=FALSE
 *   3. running (no abort, no start edge) → count if prev phase 1/2, else hold
 *
 * Counting:
 *   - Start scan: elapsed=0 (not counted)
 *   - Running scans: elapsed += 1 while prev phase 1 or 2
 *   - maxDuration: positive INT, comparison elapsed >= maxDuration triggers timeout
 *
 * Units: maxDuration in scan cycles, elapsed in scan cycles
 * Reset: Only new start rising edge (with no abort) clears elapsed/timeout
 *)

FUNCTION_BLOCK FB
VAR_INPUT
    startBtn    : BOOL;
    abortBtn    : BOOL;
    setpoint    : REAL;
    pv          : REAL;
    maxDuration : INT;
END_VAR

VAR_OUTPUT
    elapsed : INT := 0;
    phase   : INT := 0;
    timeout : BOOL := FALSE;
END_VAR

VAR
    prev_startBtn : BOOL := FALSE;
END_VAR

VAR
    startRising : BOOL;
    prev_phase  : INT;
END_VAR

// Detect rising edge of startBtn for this scan
startRising := startBtn AND NOT prev_startBtn;
prev_phase  := phase;

// Priority 1: Abort (highest)
IF abortBtn THEN
    phase := 9;
    // elapsed and timeout are preserved
    prev_startBtn := startBtn;
    RETURN;
END_IF

// Priority 2: New start rising edge (no abort)
IF startRising THEN
    phase   := 1;
    elapsed := 0;
    timeout := FALSE;
    prev_startBtn := startBtn;
    RETURN;
END_IF

// Priority 3: Running / frozen states (no abort, no new start edge)
IF prev_phase = 1 OR prev_phase = 2 THEN
    // Running: increment elapsed
    elapsed := elapsed + 1;

    IF elapsed >= maxDuration THEN
        // Timeout: enter complete state
        timeout := TRUE;
        phase   := 3;
    ELSE
        // Not yet timed out: determine phase
        IF pv >= setpoint THEN
            phase := 2;          // pv达标，保持保温
        ELSE
            phase := 1;          // 仍处于升温
        END_IF;
    END_IF;
ELSE
    // Frozen: idle (phase=0), complete (phase=3), or aborted (phase=9)
    // phase and timeout retain their values
END_IF;

prev_startBtn := startBtn;

END_FUNCTION_BLOCK

(* ---- self-hard-02.raw_candidate_03.st ---- *)
(* ENGINEERING_CONTRACT:
 * Phase activation:
 *   - Phase 0 (IDLE): Initial and idle; no counting, waiting for start
 *   - Phase 1 (HEATING): Active; elapsed increments, transitions to phase 2 on pv>=setpoint
 *   - Phase 2 (HOLDING): Active; elapsed increments, retained until timeout/abort/start
 *   - Phase 3 (COMPLETE): Retention; elapsed/timeout frozen until new start or abort
 *   - Phase 9 (ABORTED): Retention; elapsed/timeout frozen until new start
 *
 * Priority per scan (same-scan order):
 *   1. abortBtn=TRUE  → phase=9, preserve elapsed/timeout
 *   2. startBtn rising edge (no abort) → phase=1, elapsed=0, timeout=FALSE
 *   3. running (no abort, no start edge) → count if prev phase 1/2, else hold
 *
 * Counting:
 *   - Start scan: elapsed=0 (not counted)
 *   - Running scans: elapsed += 1 while prev phase 1 or 2
 *   - maxDuration: positive INT, comparison elapsed >= maxDuration triggers timeout
 *
 * Units: maxDuration in scan cycles, elapsed in scan cycles
 * Reset: Only new start rising edge (with no abort) clears elapsed/timeout
 *)

FUNCTION_BLOCK FB
VAR_INPUT
    startBtn    : BOOL;
    abortBtn    : BOOL;
    setpoint    : REAL;
    pv          : REAL;
    maxDuration : INT;
END_VAR

VAR_OUTPUT
    elapsed : INT := 0;
    phase   : INT := 0;
    timeout : BOOL := FALSE;
END_VAR

VAR
    prev_startBtn : BOOL := FALSE;
    startRising   : BOOL;
    prev_phase    : INT;
END_VAR

// Detect rising edge of startBtn for this scan
startRising := startBtn AND NOT prev_startBtn;
prev_phase  := phase;

// Priority 1: Abort (highest)
IF abortBtn THEN
    phase := 9;
    prev_startBtn := startBtn;
    RETURN;
END_IF;

// Priority 2: New start rising edge (no abort)
IF startRising THEN
    phase   := 1;
    elapsed := 0;
    timeout := FALSE;
    prev_startBtn := startBtn;
    RETURN;
END_IF;

// Priority 3: Running / frozen states (no abort, no new start edge)
IF prev_phase = 1 OR prev_phase = 2 THEN
    // Running: increment elapsed
    elapsed := elapsed + 1;

    IF elapsed >= maxDuration THEN
        // Timeout: enter complete state
        timeout := TRUE;
        phase   := 3;
    ELSE
        // Not yet timed out: determine phase
        IF pv >= setpoint THEN
            phase := 2;
        ELSE
            phase := 1;
        END_IF;
    END_IF;
END_IF;

prev_startBtn := startBtn;

END_FUNCTION_BLOCK

(* ---- self-hard-03.candidate_01.st ---- *)
(* ENGINEERING_CONTRACT
 * FIFO Queue with 8-slot compact array
 * [PUB001-PUB010] Core ops: popEn rising→remove first if count>0; pushEn rising→add pushItem if count<8
 *   Same-scan priority: pop executes BEFORE push; full→pop+push (net 0), empty→push-only (net +1)
 * [PUB011] Retention: count and fifo[1..8] state retained in VAR between scans
 * [PUB012] No AT located declarations
 * [PUB013-PUB015] Rising edge: each button triggers once per press; initial history=FALSE
 * [PUB016-PUB019] Same-scan semantics: full queue drains one slot then accepts push; empty queue accepts push only
 * [PUB020-PUB025] Array bounds: fifo[1..8], compact at end of scan: fifo[1..count] is logical queue FIFO order
 *   head=fifo[1] when non-empty, else 0; fifo[count+1..8] unspecified/unconstrained
 * [PUB026-PUB030] count∈[0,8], full↔count=8, empty↔count=0; success of push/pop updates count
 *)

(* CONTRACT_RULES [] *)

FUNCTION_BLOCK FB
VAR_INPUT
    pushEn    : BOOL;
    pushItem  : INT;
    popEn     : BOOL;
END_VAR
VAR_IN_OUT
    fifo      : ARRAY[1..8] OF INT;
END_VAR
VAR_OUTPUT
    count     : INT;
    full      : BOOL;
    empty     : BOOL;
    head      : INT;
END_VAR
VAR
    prev_pushEn : BOOL := FALSE;
    prev_popEn  : BOOL := FALSE;
    tmp_pushRising : BOOL;
    tmp_popRising  : BOOL;
    tmp_i       : INT;
END_VAR

    // Rising edge detection
    tmp_popRising  := popEn AND NOT prev_popEn;
    tmp_pushRising := pushEn AND NOT prev_pushEn;
    prev_popEn  := popEn;
    prev_pushEn := pushEn;

    // Execute in required order: pop first, then push
    // POP: non-empty queue only
    IF tmp_popRising AND count > 0 THEN
        FOR tmp_i := 1 TO count - 1 DO
            fifo[tmp_i] := fifo[tmp_i + 1];
        END_FOR;
        count := count - 1;
    END_IF;

    // PUSH: non-full queue only
    IF tmp_pushRising AND count < 8 THEN
        count := count + 1;
        fifo[count] := pushItem;
    END_IF;

    // Outputs
    full  := (count = 8);
    empty := (count = 0);
    IF empty THEN
        head := 0;
    ELSE
        head := fifo[1];
    END_IF;

END_FUNCTION_BLOCK
